(* IEC 61131-3 sources: daoli-st-library/DL_Algo (part 3) *)

(* ---- FB_DL_ThermalRampPredict.st ---- *)
(*==============================================================================
 * 组件名称 (Component)  : FB_DL_ThermalRampPredict
 * 所属子库 (Sublibrary) : DL_Algo
 * 当前版本 (Version)    : 1.0.0
 * 兼容性   (Platform)   : CODESYS 3.5+ / TwinCAT 3 / 汇川 InoProShop / 施耐德 Machine Expert
 *                         仅依赖 Standard.library（R_TRIG / ABS / MIN / MAX）与库内时间换算内核
 *                         FC_DL_TimeToLrealSec / FC_DL_LrealSecToTime，零厂商私有库
 * 功能描述 (Function)   : 一阶热模型预测与前馈。模型 dT/dt = 〔u·K − (T − Tamb)〕/ tau，本件不驱 u，
 *                         而以「满功率模型斜率」作参考，用实测斜率在线修正时间常数 tau：
 *                         ① tRemain：据当前温度、目标温度与实测斜率外推到目标所需剩余时间；
 *                         ② fFfBias：进入目标前 fLeadBand 带内按接近程度线性加大「减功率量」，
 *                         抑制热惯性造成的超调（前馈偏移，非闭环）；
 *                         ③ tau 在线修正：实测斜率与模型斜率偏差持续超阈值时按 ±5% 微调，
 *                         并钳在〔tTauMin, tTauMax〕，防单次扰动把模型带偏。
 * 分工声明 (Scope)      : 与 `FB_DL_DryingOvenZone` / `FB_DL_CvdTempRamp`（分区控温与温度曲线
 *                         执行）分工 —— 本件**只出预测与前馈偏置**，不闭环、不持曲线、不下发
 *                         加热指令；曲线执行与闭环属主为上列两件。
 * 接口     (Interface)  : 输入 fTempC 当前温度、fTargetC 目标温度、fAmbC 环境温度、fGainK 稳态
 *                         增益、tTau 时间常数、tTauMin / tTauMax 修正上下限、fLeadBand 前馈起始带、
 *                         fFfBiasMax 前馈偏置上限、fSlopeDevMax 斜率偏差阈值、tTaskPeriod 任务周期、
 *                         bEnable 使能、bReset 复位；输出 tRemain 剩余时间（无趋势时为哨兵）、
 *                         bNoTrend 无趋势标志、fFfBias 前馈减功率量、fTauUsed 当前使用的时间常数、
 *                         eState / eCause / bError / nErrId。
 * 边界     (Boundary)   : ① 组态闸：tTau <= T#0S、tTauMin <= T#0S、tTauMax <= tTauMin、fGainK <= 0.0、
 *                         fLeadBand <= 0.0、fFfBiasMax <= 0.0、fSlopeDevMax < 0.0、tTaskPeriod <= T#0S
 *                         或任一浮点引脚 NaN → 故障锁存（每个参与判据的引脚都在闸内，R151）；
 *                         ② tRemain 计算防除零：当实测斜率绝对值 <= DL_SLOPE_EPS 时**不返回 T#0S**
 *                         （T#0S 会被上层读成「马上就到」），而返回哨兵 DL_TIME_INF 并置 bNoTrend；
 *                         ③ 前馈偏置双侧钳位〔0.0, fFfBiasMax〕，禁单侧钳位；
 *                         ④ 非有限输入 → 故障闸，输出侧 tRemain 哨兵、fFfBias 0（安全侧）；
 *                         ⑤ R_TRIG 一枚段 0 无条件周期刷新；⑥ 故障相迁出唯一路径 = bReset 上升沿；
 *                         ⑦ 零全局耦合（无 GVL / 无物理地址）。
 * 遗留假设 (Assumption) : 【R95 三句声明】① 代理值 = 引脚 tTaskPeriod，用于把逐拍温差换算成 °C/s；
 *                         ② 覆盖范围 = 任务周期 10 ms ~ 2 s 的周期任务；③ 覆盖不到的区间
 *                         （< 10 ms 的高速任务或超载抖动任务）由调用方负责：此时斜率噪声偏大，
 *                         tau 修正应经 bEnable 关断，仅使用 fFfBias 前馈。
 * 解除式   (Release)    : bReset 上升沿 ∧ 组态合法 ∧ 非无趋势（NOT bNoTrend，当拍量）。
 *                         自证可满足（终审两式 1）：bNoTrend 由当拍斜率派生，温度一旦真实变化
 *                         斜率即非零，标志必落假；解除式不含计时器输出与锁存量比较，无恒假因子。
 * 码表     (Codes)      : 16#0002_03B3 故障级：热模型预测故障总码（组态非法 / 输入非有限 / 非法
 *                         相位），锁存至 bReset 上升沿，归因由 eCause 承载（R190 单件单总码）；
 *                         16#0002_04B6 信息级：无趋势（斜率近似为 0，剩余时间输出哨兵）。
 *                         加码反证（R90）：无趋势时 tRemain 是哨兵常量、fFfBias 仍有效，若只靠
 *                         「tRemain = 86400 s」判断，上层无法区分「真的还要一天」与「算不出来」，
 *                         故须立一码（bNoTrend 只是布尔位，不进报警台账）。
 *                         码段说明：0002 段故障子带 03xx / 信息子带 04xx，本件取 03B3 / 04B6
 *                         （源码实扫该两槽为空，续接同子带已用最大值，未回填碎片孔洞）。
 * 编译门槛 (Build Gate) : 本件委托 FC_DL_TimeToLrealSec 与 FC_DL_LrealSecToTime（内部转调平台
 *                         内建 TIME_TO_LREAL / LREAL_TO_TIME），交付门槛：须在 CODESYS / TwinCAT 3 /
 *                         InoProShop 三平台各编译验证一次。
 * 开源溯源 (Origin)     : 道莅自研 clean-room（参考一阶热模型与时间常数在线修正参数域，
 *                         零代码行复制；t2-1-lgf 技术子族）
 * 修订历史 (Revision)   : 2026-11-19  v1.0.0  R45 首版（批次 2 · 序号 9）
 *==============================================================================*)

TYPE E_DL_TrpState :
(
    eIdle  := 0,     // 失能待使能 / Idle, disabled
    eRun   := 10,    // 预测运行 / Predicting in run
    eFault := 90     // 故障锁存相 / Fault latched phase
);
END_TYPE

TYPE E_DL_TrpCause :
(
    eNone       := 0,   // 无故障成因 / No cause
    eCfgIllegal := 1,   // 组态非法 / Illegal configuration
    eNonFinite  := 2,   // 输入非有限 / Non-finite input
    ePhaseBad   := 3    // 非法相位兜底 / Illegal phase fallback
);
END_TYPE

FUNCTION_BLOCK FB_DL_ThermalRampPredict
VAR_INPUT
    fTempC        : REAL := 25.0;       // 当前温度 [°C] / Current temperature [degC]
    fTargetC      : REAL := 80.0;       // 目标温度 [°C] / Target temperature [degC]
    fAmbC         : REAL := 25.0;       // 环境温度 [°C] / Ambient temperature [degC]
    fGainK        : REAL := 55.0;       // 稳态增益（满功率温升上界），域 > 0.0 [°C] / Steady-state gain, domain > 0.0 [degC]
    tTau          : TIME := T#120S;     // 时间常数初值，域 > T#0S [ms] / Initial time constant, domain > T#0S [ms]
    tTauMin       : TIME := T#20S;      // 修正下限，域 > T#0S 且 < tTauMax [ms] / Correction lower bound [ms]
    tTauMax       : TIME := T#900S;     // 修正上限，域 > tTauMin [ms] / Correction upper bound [ms]
    fLeadBand     : REAL := 10.0;       // 前馈起始带（距目标多近开始减功率），域 > 0.0 [°C] / Lead band, domain > 0.0 [degC]
    fFfBiasMax    : REAL := 60.0;       // 前馈减功率量上限，域 > 0.0 [%] / Feed-forward bias ceiling, domain > 0.0 [%]
    fSlopeDevMax  : REAL := 0.05;       // 斜率偏差阈值（相对值），域 >= 0.0 [p.u.] / Slope deviation threshold [p.u.]
    tTaskPeriod   : TIME := T#100MS;    // 调用任务周期（代理值，见头注释遗留假设），域 > T#0S [ms] / Task period proxy [ms]
    bEnable       : BOOL := TRUE;       // 预测使能 [-] / Prediction enable
    bReset        : BOOL := FALSE;      // 复位命令，上升沿清故障 [-] / Reset command, rising edge clears fault
END_VAR
VAR_OUTPUT
    tRemain       : TIME;               // 剩余时间（无趋势时输出哨兵 24 h） [ms] / Remaining time, sentinel 24 h when no trend [ms]
    bNoTrend      : BOOL;               // 无趋势标志（斜率近似 0） [-] / No-trend flag
    fFfBias       : REAL;               // 前馈减功率量（双侧钳位后） [%] / Feed-forward power reduction, clamped [%]
    fTauUsed      : REAL;               // 当前使用的时间常数（在线修正后） [s] / Time constant in use after correction [s]
    eState        : E_DL_TrpState;      // 状态出口，段 6 单点映射 / State outlet
    eCause        : E_DL_TrpCause;      // 故障成因出口（R190 归因唯一） / Fault cause outlet
    bError        : BOOL;               // 故障锁存标志 [-] / Fault latch flag
    nErrId        : UDINT;              // 事件码，0 = 无事件 / Event code, 0 = no event
END_VAR
VAR
    _eState       : E_DL_TrpState := E_DL_TrpState.eIdle;   // 内部相位（CASE 唯一写入目标） / Internal phase
    _eCause       : E_DL_TrpCause := E_DL_TrpCause.eNone;   // 故障成因锁存（锁存量） / Latched cause
    rtReset       : R_TRIG;             // 复位沿实例，段 0 无条件调用 / Reset edge
    _fTsSec       : LREAL;              // 任务周期秒数（当拍量） [s] / Task period in seconds
    _fTauSec      : LREAL;              // 时间常数秒数（当拍量，取自修正后的 tTau） [s] / Time constant in seconds
    _fTempPrev    : REAL;               // 上拍温度快照（锁存量） [°C] / Previous-scan temperature snapshot
    _fSlopeMeas   : LREAL;              // 实测斜率（当拍量） [°C/s] / Measured slope [degC/s]
    _fSlopeModel  : LREAL;              // 满功率模型斜率（当拍量） [°C/s] / Full-power model slope [degC/s]
    _fDeltaT      : REAL;               // 目标 − 当前温差 [°C] / Target minus current temperature [degC]
    _fRemSec      : LREAL;              // 剩余时间秒数（转换前） [s] / Remaining seconds before conversion
    _fTauUsedSec  : LREAL;              // 在线修正后的时间常数（锁存量） [s] / Corrected time constant, latched
    _nDevRun      : INT;                // 斜率偏差持续计数（锁存量） [拍] / Slope deviation persistence counter, latched
    _uConvErrT    : UDINT;              // 周期换算错误码（当拍量） [-] / Period conversion error code
    _uConvErrU    : UDINT;              // 时间常数换算错误码（当拍量） [-] / Tau conversion error code
    _uConvErrR    : UDINT;              // 剩余时间换算错误码（当拍量） [-] / Remaining-time conversion error code
    _bConvErrT    : BOOL;               // 周期换算故障位（当拍量） [-] / Period conversion fault flag
    _bConvErrU    : BOOL;               // 时间常数换算故障位（当拍量） [-] / Tau conversion fault flag
    _bConvErrR    : BOOL;               // 剩余时间换算故障位（当拍量） [-] / Remaining-time conversion fault flag
    _bConvValidT  : BOOL;               // 周期换算有效位（当拍量） [-] / Period conversion valid flag
    _bConvValidU  : BOOL;               // 时间常数换算有效位（当拍量） [-] / Tau conversion valid flag
    _bConvValidR  : BOOL;               // 剩余时间换算有效位（当拍量） [-] / Remaining-time conversion valid flag
    _bInit        : BOOL;               // 首拍初始化完成位（锁存量） [-] / First-scan init done
    _bNonFin      : BOOL;               // 输入非有限当拍量 [-] / Non-finite input this scan
    _bCfgBad      : BOOL;               // 组态非法当拍量 [-] / Illegal configuration
    _bFault       : BOOL;               // 故障锁存位（锁存量） / Latched fault bit
    _uFault       : UDINT;              // 故障码锁存（锁存量） / Latched fault code
    _uInfo        : UDINT;              // 信息码，每拍重算 / Info code, recomputed each scan
END_VAR
VAR CONSTANT
    DL_FLOAT_EPS  : LREAL := 1.0E-6;    // 浮点判零容差 [无量纲] / Float epsilon for zero tests
    DL_SLOPE_EPS  : LREAL := 1.0E-4;    // 斜率判零容差（低于此判无趋势） [°C/s] / Slope epsilon, below means no trend [degC/s]
    DL_TIME_INF   : LREAL := 86400.0;   // 「无趋势」哨兵秒数（24 h，远离任何真实剩余时间） [s] / No-trend sentinel seconds, 24 h [s]
    DL_TAU_STEP   : LREAL := 1.05;      // 时间常数单次修正倍率 [-] / Time constant correction factor per adjustment
    DL_DEV_MAX    : INT := 10;          // 斜率偏差持续拍数门限 [拍] / Slope deviation persistence limit [scan]
END_VAR

(* —— 段 0：当拍判据派生 + 沿实例无条件周期刷新 —— *)
_fTsSec := FC_DL_TimeToLrealSec(tIn := tTaskPeriod, eErr => _uConvErrT, bError => _bConvErrT, bValid => _bConvValidT);   // 周期换算（R140 委托） / Period conversion
_fTauSec := FC_DL_TimeToLrealSec(tIn := tTau, eErr => _uConvErrU, bError => _bConvErrU, bValid => _bConvValidU);         // 时间常数换算 / Tau conversion
_bNonFin := (fTempC <> fTempC) OR (fTargetC <> fTargetC) OR (fAmbC <> fAmbC) OR (fGainK <> fGainK)    // NaN 自反判（判等禁令唯一例外） / NaN self-reflexive tests
         OR (fLeadBand <> fLeadBand) OR (fFfBiasMax <> fFfBiasMax) OR (fSlopeDevMax <> fSlopeDevMax); // 前馈参数 NaN 判 / Feed-forward parameter NaN tests
_bCfgBad := (tTau <= T#0S) OR (tTauMin <= T#0S) OR (tTauMax <= tTauMin) OR (tTaskPeriod <= T#0S)     // 时间类组态闸 / Time config gates
            OR (fGainK <= 0.0) OR (fLeadBand <= 0.0) OR (fFfBiasMax <= 0.0) OR (fSlopeDevMax < 0.0)   // 浮点域闸（R151 全覆盖） / Float domain gates
            OR (_uConvErrT <> 16#0000_0000) OR (_uConvErrU <> 16#0000_0000);                          // 换算错误并入闸 / Conversion errors folded in
rtReset(CLK := bReset);                                                                              // 复位沿，每拍必调（R228A） / Reset edge

(* —— 段 1：单拍量预清零（锁存量与快照量不入清单，R107） —— *)
_uInfo   := 16#0000_0000;          // 信息码每拍重算 / Info recomputed every scan
bNoTrend := FALSE;                 // 无趋势标志每拍预清 / No-trend flag preset
nErrId   := 16#0000_0000;          // 事件码缺省无事件 / Event code default none
bError   := FALSE;                 // 故障标志每拍预清，故障分支同拍置位（R45 配对） / Flag preset
fFfBias  := 0.0;                   // 前馈偏置缺省 0（安全侧：不减功率） / Bias default 0, safe side

(* —— 段 2：复位沿 + 组态域闸 + 非有限闸 —— *)
IF rtReset.Q THEN                                                        // 当拍复位沿 / current-scan reset edge
    _bFault := FALSE;                                                    // 清故障锁存位（锁存量） / Clear fault latch
    _uFault := 16#0000_0000;                                             // 清故障锁存码（锁存量） / Clear latched code
    _eCause := E_DL_TrpCause.eNone;                                      // 清成因（锁存量） / Clear latched cause
    IF _eState = E_DL_TrpState.eFault THEN
        _eState := E_DL_TrpState.eIdle;                                  // 故障相迁出唯一路径 / Sole exit from fault phase
    END_IF
END_IF
IF _bCfgBad THEN                                                         // 组态域闸 / Configuration gate
    _uFault := 16#0002_03B3;                                             // 故障级：热模型预测故障总码 / Fault-level: prediction fault code
    _bFault := TRUE;
    bError  := TRUE;                                                     // 故障标志同拍置位（R45 配对） / Error flag set same scan
    _eCause := E_DL_TrpCause.eCfgIllegal;                                // 归因：组态非法 / Cause: illegal configuration
END_IF
IF (NOT _bFault) AND _bNonFin THEN                                       // 输入非有限 / Non-finite input
    _uFault := 16#0002_03B3;
    _bFault := TRUE;
    bError  := TRUE;
    _eCause := E_DL_TrpCause.eNonFinite;                                 // 归因：非有限 / Cause: non-finite
END_IF

(* —— 段 3：时间常数初始化（首拍取初值并钳在修正域内） —— *)
IF NOT _bInit THEN
    IF _fTauSec < FC_DL_TimeToLrealSec(tIn := tTauMin) THEN              // 初值低于下限即钳入域内 / Clamp initial value into domain
        _fTauUsedSec := FC_DL_TimeToLrealSec(tIn := tTauMin);
    ELSIF _fTauSec > FC_DL_TimeToLrealSec(tIn := tTauMax) THEN
        _fTauUsedSec := FC_DL_TimeToLrealSec(tIn := tTauMax);
    ELSE
        _fTauUsedSec := _fTauSec;
    END_IF
    _fTempPrev := fTempC;                                                // 温度快照初始化 / Initialize temperature snapshot
    _bInit := TRUE;                                                      // 初始化完成 / Init done
END_IF

(* —— 段 4：斜率测量、模型斜率与时间常数在线修正（仅无故障且使能） —— *)
IF (NOT _bFault) AND bEnable THEN
    IF _fTsSec > DL_FLOAT_EPS THEN                                       // 除零前置判 / Divide-by-zero guard
        _fSlopeMeas := REAL_TO_LREAL(fTempC - _fTempPrev) / _fTsSec;      // 实测斜率 [°C/s] / Measured slope
    ELSE
        _fSlopeMeas := 0.0;                                              // 周期退化时置 0（组态闸已拦，防御纵深） / Degenerate period
    END_IF
    IF _fTauUsedSec > DL_FLOAT_EPS THEN                                  // 除零前置判 / Divide-by-zero guard
        _fSlopeModel := REAL_TO_LREAL(fGainK - (fTempC - fAmbC)) / _fTauUsedSec;   // 满功率模型斜率 / Full-power model slope
    ELSE
        _fSlopeModel := 0.0;                                             // 退化兜底 / Degenerate guard
    END_IF
    IF ABS(_fSlopeModel) > DL_SLOPE_EPS THEN                             // 相对偏差需有非零参照 / Relative deviation needs a non-zero reference
        IF ABS((_fSlopeMeas - _fSlopeModel) / _fSlopeModel) > fSlopeDevMax THEN
            IF _nDevRun < DL_DEV_MAX THEN
                _nDevRun := _nDevRun + 1;                                // 偏差持续计数 / Deviation persistence count
            END_IF
        ELSE
            _nDevRun := 0;                                               // 回到阈值内即清零 / Reset inside threshold
        END_IF
    ELSE
        _nDevRun := 0;
    END_IF
    IF _nDevRun >= DL_DEV_MAX THEN                                       // 偏差持续：按符号微调时间常数 / Sustained deviation, adjust tau by sign
        IF _fSlopeMeas < _fSlopeModel THEN                               // 实测偏慢 → 时间常数变大 / Slower than model, tau up
            _fTauUsedSec := MIN(_fTauUsedSec * DL_TAU_STEP, FC_DL_TimeToLrealSec(tIn := tTauMax));
        ELSE
            _fTauUsedSec := MAX(_fTauUsedSec / DL_TAU_STEP, FC_DL_TimeToLrealSec(tIn := tTauMin));
        END_IF
        _nDevRun := 0;                                                   // 修正后计数清零 / Reset after correction
    END_IF
END_IF

(* —— 段 5：剩余时间预测（防除零；无趋势输出哨兵而非 T#0S） —— *)
IF (NOT _bFault) AND bEnable THEN
    _fDeltaT := fTargetC - fTempC;                                       // 剩余温差 / Remaining temperature difference
    IF ABS(_fSlopeMeas) <= DL_SLOPE_EPS THEN                             // 斜率近似 0：不得输出 T#0S 冒充「马上到」 / Slope near zero, never emit T#0S
        bNoTrend := TRUE;                                                // 无趋势标志 / No-trend flag
        _fRemSec := DL_TIME_INF;                                         // 哨兵秒数 / Sentinel seconds
        _uInfo := 16#0002_04B6;                                          // 信息级：无趋势留痕 / Info: no trend recorded
    ELSE
        _fRemSec := REAL_TO_LREAL(_fDeltaT) / _fSlopeMeas;               // 线性外推剩余时间 / Linear extrapolation
        IF _fRemSec < 0.0 THEN                                           // 已越过目标（过冲在恢复）：剩余判 0 而非负数 / Already past target
            _fRemSec := 0.0;
        END_IF
        IF _fRemSec > DL_TIME_INF THEN                                   // 上界兜底防 TIME 溢出 / Upper bound guard
            _fRemSec := DL_TIME_INF;
        END_IF
    END_IF
    tRemain := FC_DL_LrealSecToTime(fSec := _fRemSec, eErr => _uConvErrR, bError => _bConvErrR, bValid => _bConvValidR);   // 委托时间换算 / Delegate conversion
ELSE
    tRemain := FC_DL_LrealSecToTime(fSec := DL_TIME_INF);                // 非运行相输出哨兵（不宣称「马上到」） / Sentinel outside run phase
END_IF

(* —— 段 6：前馈偏置（进入 fLeadBand 带内线性加大减功率量，双侧钳位） —— *)
IF (NOT _bFault) AND bEnable THEN
    IF ABS(_fDeltaT) < fLeadBand THEN                                    // 进入前馈带 / Inside lead band
        fFfBias := fFfBiasMax * (1.0 - (ABS(_fDeltaT) / fLeadBand));      // 越接近目标减得越多 / More reduction as target nears
    ELSE
        fFfBias := 0.0;                                                  // 带外不减功率 / No reduction outside band
    END_IF
    IF fFfBias > fFfBiasMax THEN                                         // 双侧钳位（上侧） / Two-sided clamp, upper
        fFfBias := fFfBiasMax;
    END_IF
    IF fFfBias < 0.0 THEN                                                // 双侧钳位（下侧） / Two-sided clamp, lower
        fFfBias := 0.0;
    END_IF
END_IF

(* —— 段 7：温度快照更新（主体末行，跨拍纪律） —— *)
_fTempPrev := fTempC;                                                    // 温度快照（本拍末更新） / Temperature snapshot at body end

(* —— 段 8：故障解除式（R240 全当拍量） —— *)
IF rtReset.Q AND (NOT _bCfgBad) AND (NOT _bNonFin) AND (NOT bNoTrend) THEN
    _bFault := FALSE;                                                    // 清故障锁存位（锁存量） / Clear fault latch
    _uFault := 16#0000_0000;                                             // 清故障锁存码（锁存量） / Clear latched code
    _eCause := E_DL_TrpCause.eNone;                                      // 清成因（锁存量） / Clear latched cause
END_IF

(* —— 段 8A：故障锁存相位迁移闸 —— *)
IF _bFault AND (_eState <> E_DL_TrpState.eFault) THEN
    _eState := E_DL_TrpState.eFault;                                     // 锁存即入故障相 / Latch enters fault phase
END_IF

(* —— 段 9：相位机（ENUM 全成员显式标签 + ELSE 兜底，R128） —— *)
CASE _eState OF

E_DL_TrpState.eIdle:
    IF bEnable AND _bInit AND (NOT _bFault) THEN                         // 出口 1：使能且已初始化 / Enabled and initialized
        _eState := E_DL_TrpState.eRun;
    ELSIF _bFault THEN                                                   // 出口 2：故障锁存 / Fault latched
        _eState := E_DL_TrpState.eFault;
    END_IF

E_DL_TrpState.eRun:
    IF (NOT bEnable) THEN                                                // 出口 1：失能（前置消失，R98） / Disabled
        _eState := E_DL_TrpState.eIdle;
    ELSIF _bFault THEN                                                   // 出口 2：故障锁存 / Fault latched
        _eState := E_DL_TrpState.eFault;
    END_IF

E_DL_TrpState.eFault:
    ;                                                                     // 故障相：仅段 8 复位沿可迁出 / Only the reset edge leaves this phase

ELSE
    _uFault := 16#0002_03B3;                                             // 故障级：非法相位兜底（归并总码） / Illegal-phase fallback
    _bFault := TRUE;
    bError  := TRUE;
    _eCause := E_DL_TrpCause.ePhaseBad;                                  // 归因：非法相位 / Cause: illegal phase
    _eState := E_DL_TrpState.eFault;

END_CASE

(* —— 段 10：出口单点映射（名实同源；锁存码回放；故障相安全侧） —— *)
IF _bFault THEN
    tRemain  := FC_DL_LrealSecToTime(fSec := DL_TIME_INF);               // 故障相输出哨兵（不宣称短时到达） / Sentinel in fault
    bNoTrend := TRUE;                                                    // 故障相判无趋势（不给出时间承诺） / No-trend in fault
    fFfBias  := 0.0;                                                     // 故障相不减功率（不加未知偏置） / No bias in fault
    fTauUsed := LREAL_TO_REAL(_fTauUsedSec);                             // 时间常数镜像（供调试） / Tau mirror for commissioning
ELSIF NOT bEnable THEN
    fTauUsed := LREAL_TO_REAL(_fTauUsedSec);                             // 失能相仍回放时间常数（观测语义） / Tau echoed when disabled
    tRemain  := FC_DL_LrealSecToTime(fSec := DL_TIME_INF);               // 失能相哨兵 / Sentinel when disabled
    bNoTrend := TRUE;                                                    // 失能相无预测 / No prediction when disabled
ELSE
    fTauUsed := LREAL_TO_REAL(_fTauUsedSec);                             // 运行相时间常数 / Tau in run
END_IF
IF _bFault THEN
    nErrId := _uFault;                                                   // 故障锁存码回放 / Replay latched fault code
ELSE
    nErrId := _uInfo;                                                    // 信息码 / Info code
END_IF
bError := _bFault;                                                       // 故障标志与锁存同源（名实双出口，R191） / Flag from latch
eState := _eState;                                                       // 状态出口 / State outlet
eCause := _eCause;                                                       // 成因出口 / Cause outlet

END_FUNCTION_BLOCK

(* ---- FB_DL_ValveCharacteristic.st ---- *)
(*==============================================================================
 * 组件名称 (Component)  : FB_DL_ValveCharacteristic
 * 所属子库 (Sublibrary) : DL_Algo
 * 当前版本 (Version)    : 1.0.1
 * 兼容性   (Platform)   : CODESYS 3.5 / TwinCAT 3 / 汇川 InoProShop / Machine Expert
 *                         仅依赖 Standard.library（ABS / LN / SQRT / MIN / MAX / R_TRIG）
 * 功能描述 (Function)   : 把「期望流量百分比」按调节阀固有特性折算为「阀位百分比」，
 *                         支持线性 / 等百分比 / 快开三种特性，带可调比、行程上下限、
 *                         输出死区与饱和标志。现场用途：等百分比阀按线性给定会让小流量段
 *                         分辨率不足、大流量段增益过高并引起振荡；本件把特性补偿收回
 *                         PLC 侧，工艺员不再靠「凭经验把给定调弯」。
 *                         死区只压输出抖动，不改变内部限幅结果；掉使能保持上次阀位
 *                         （阀位突跳比保持更危险），阀位回零由上层安全逻辑负责。
 * 出口契约 (Exit)       : fTravel 为最终阀位给定，域为生效行程上下限之间；
 *                         bSaturated 表示输出被流量给定域、可调比下限或行程上下限任一截断；
 *                         bError 为故障级锁存，只由 2010 / 2011 / 2012 三码置位，
 *                         bReset 上升沿清故障回空闲。信息码 2001 / 2002 / 2003 每拍重算。
 * 开源溯源 (Origin)     : 来源标签 isa88-process（工艺参数域）。许可证：ISA-88 为公开标准，
 *                         无源码可复制；调节阀流量特性公式取自公开的过程控制教材定义。
 *                         借鉴点：把「特性」做成**枚举参数域**而非三个独立功能块——三种特性
 *                         共用同一套限幅、死区与状态机，拆块会产生三份重复代码，
 *                         且特性切换在配方里属于运行期行为。
 *                         clean-room 独立实现，与任何厂商阀门功能块无代码关联。
 * 码位说明 (Codes)      : 信息级 16#0002_2001（输出被下限截断）/ 2002（输出被上限截断）/
 *                         2003（死区保持）；故障级 16#0002_2010（行程配置非法）/
 *                         2011（可调比对数的二次守卫触发）/ 2012（非法特性枚举兜底）。
 *                         共 6 码，全部落在 R12 计划第 1.2 节本件码段内。
 * 依赖     (Depends)    : 无 DL_ 内部依赖；Standard.library: ABS / LN / SQRT / MAX / R_TRIG
 * 红线自检 (Redline)    : 1 ✓ 零全局变量表依赖、零外部变量声明、零物理地址
 *                         2 ✓ 纯 IEC 61131-3，无指针、无厂商库
 *                         3 ✓ 对数与开方先做域守护、可调比下限保证对数分母不为零、
 *                             行程上下限倒置直接判故障而不交换、死区比较用容差不用判等
 *                         4 ✓ 全变量中英双语同行注释
 *                         5 ✓ 三态 ENUM + CASE 全覆盖 + ELSE 兜底（2012）；特性选择亦全覆盖
 *                         6 ✓ R_TRIG 实例在 CASE 之外每拍无条件刷新
 *                         7 ✓ END_FUNCTION_BLOCK 位于文件最后有效行
 * 规格偏离留档 (Deviation):
 *   计划 3.11 节正文提到 2004 / 2005 / 2006 三个「输入钳位」码，但同计划第 1.2 节给本件
 *   只分配了 2001~2003 与 2010~2012 六个码，两者冲突。按「码位表为准、不得自创」的纪律，
 *   本实现对输入钳位采取如下归并：流量给定越界钳位并入 2001 / 2002（越界必然让输出打端点，
 *   语义与截断一致）；可调比与死区的钳位属整定参数修正，不单独置码，仅钳位后照算，
 *   并在头注释与本段注释中写明，不再占用段外码。
 * 修订历史 (Revision)   :
 *   2026-11-15  v1.0.0  首版入库（R12 · DL_Algo 工艺参数域）
 *   2026-11-15  v1.0.1  终审修复：投运与故障复位首拍不再强制阀位回行程下限
 *                       （原实现 fLast := fLoTravel 会让阀门在复位当拍直冲最小开度，
 *                       与本件「不做阀位回零、突跳比保持更危险」的契约自相矛盾）；
 *                       改为「保持上次阀位并夹到生效行程内」，同时补齐行程域的出口保证
 *============================================================================*)

(*-----------------------------------------------------------------------------
 * 枚举: E_DL_ValveCharKind（归属 DL_Algo，与本功能块同文件）
 * 含义: 调节阀固有流量特性。三种特性共用同一套限幅与死区逻辑。
 *----------------------------------------------------------------------------*)
TYPE E_DL_ValveCharKind :
(
    eLinear       := 0,    // 线性特性：阀位与流量成正比 / Linear: travel proportional to flow
    eEqualPercent := 10,   // 等百分比特性：单位阀位变化引起的流量变化与当前流量成正比 / Equal percentage
    eQuickOpen    := 20    // 快开特性：小阀位即获大流量，后段渐平 / Quick opening, fast rise then flat
);
END_TYPE

(*-----------------------------------------------------------------------------
 * 枚举: E_DL_ValveCharState（归属 DL_Algo，与本功能块同文件）
 * 含义: 特性补偿块的离散状态。
 *----------------------------------------------------------------------------*)
TYPE E_DL_ValveCharState :
(
    eIdle   := 0,     // 空闲：等待使能与行程配置校验 / Idle: waiting for enable and travel validation
    eActive := 10,    // 运行：折算特性、限幅、死区、输出 / Active: convert, clamp, deadband, publish
    eFault  := 99     // 故障：配置非法或枚举兜底，输出保持上次 / Fault: invalid config, travel held
);
END_TYPE

(*==============================================================================
 * 功能块: FB_DL_ValveCharacteristic
 * 调用约定: 每个扫描周期无条件调用一次；bEnable 为 FALSE 时阀位保持上次值。
 * 无状态泄漏: 全部状态驻留于实例私有 VAR，零全局引用，可多实例并行。
 *============================================================================*)
FUNCTION_BLOCK FB_DL_ValveCharacteristic
VAR_INPUT
    bEnable       : BOOL;                                // 使能，FALSE 时阀位保持上次输出 / Enable, holds the last travel when FALSE
    bReset        : BOOL;                                // 上升沿清故障回空闲 / Rising edge clears the fault
    fFlowCmd      : REAL := 0.0;                         // 期望流量 [百分比]，域 0~100 / Desired flow in percent, 0..100
    eChar         : E_DL_ValveCharKind := E_DL_ValveCharKind.eEqualPercent;  // 固有特性 [-] / Inherent characteristic
    fRangeability : REAL := 30.0;                        // 可调比 [-]，域 2~100，越界钳位 / Rangeability, clamped to 2..100
    fMinTravel    : REAL := 0.0;                         // 最小阀位 [百分比]，域 0~100 / Minimum travel in percent
    fMaxTravel    : REAL := 100.0;                       // 最大阀位 [百分比]，域 0~100 / Maximum travel in percent
    fDeadband     : REAL := 0.2;                         // 输出死区 [百分比]，变化小于此值保持上次 / Output deadband in percent
END_VAR
VAR_OUTPUT
    fTravel       : REAL;                                // 阀位给定 [百分比]，域 fMinTravel~fMaxTravel / Travel command in percent
    bSaturated    : BOOL;                                // 输出被上下限或可调比下限截断 TRUE / Output clamped
    bError        : BOOL;                                // 故障级锁存，仅 2010~2012 置位 / Latched fault
    uErrorId      : UDINT;                               // 事件码，0 = 无事件 / Event code, zero means none
    eState        : E_DL_ValveCharState;                 // 主状态机当前状态 / Current state
END_VAR
VAR
    fbTrigReset   : R_TRIG;                              // 复位沿，CASE 之外每拍刷新 / Reset edge, refreshed outside CASE
    ePhase        : E_DL_ValveCharState := E_DL_ValveCharState.eIdle;  // 内部状态 / Internal state
    fFlowVal      : REAL;                                // 钳位后的期望流量 [百分比] / Clamped flow command in percent
    fQ            : REAL;                                // 归一化流量 [0~1] / Normalised flow
    fR            : REAL;                                // 生效可调比 [-] / Effective rangeability
    fRaw          : REAL;                                // 未限幅的阀位 [百分比] / Unlimited travel in percent
    fLast         : REAL;                                // 上次输出阀位 [百分比] / Last travel command
    fLoTravel     : REAL;                                // 生效行程下限 [百分比] / Effective lower bound
    fHiTravel     : REAL;                                // 生效行程上限 [百分比] / Effective upper bound
    fQMin         : REAL;                                // 可调比下限对应的归一化流量 [0~1] / Normalised flow at the rangeability floor
    fDeadUse      : REAL;                                // 生效死区宽度 [百分比] / Effective deadband width
    bClampLo      : BOOL;                                // 下限截断标记 / Lower clamp flag
    bClampHi      : BOOL;                                // 上限截断标记 / Upper clamp flag
END_VAR
VAR CONSTANT
    DL_PCT_MAX    : REAL := 100.0;                       // 百分比满量程 [百分比] / Percent full scale
    DL_R_MIN      : REAL := 2.0;                         // 可调比下限 [-] / Minimum rangeability
    DL_R_MAX      : REAL := 100.0;                       // 可调比上限 [-] / Maximum rangeability
    DL_DB_MAX     : REAL := 5.0;                         // 死区宽度上限 [百分比] / Deadband ceiling in percent
    DL_EPS        : REAL := 1.0E-6;                      // 浮点判零容差 [-] / Float zero tolerance
END_VAR

(*------------------------------------------------------------------------------
 * 段 1｜复位沿每拍无条件刷新（严禁放进 CASE 内部）
 *      Reset edge refreshed unconditionally on every scan
 *-----------------------------------------------------------------------------*)
fbTrigReset(CLK := bReset);

(*------------------------------------------------------------------------------
 * 段 2｜输入调理：流量给定的域钳位，与整定参数的可调比 / 死区钳位
 *      Input conditioning: flow clamp plus rangeability and deadband clamps
 *      流量越界钳位必然把输出打到端点，语义等同截断，故并入 2001 / 2002 报码
 *      A clamped flow command drives the output to an end point, reported as 2001 / 2002
 *      可调比与死区的钳位只是整定参数修正，不单独置码，钳位后照算
 *      Rangeability and deadband clamps are tuning fixes and carry no dedicated code
 *-----------------------------------------------------------------------------*)
bClampLo  := FALSE;
bClampHi  := FALSE;
fFlowVal  := fFlowCmd;
IF NOT (fFlowVal >= 0.0) THEN
    fFlowVal := 0.0;
    bClampLo := TRUE;
ELSIF fFlowVal > DL_PCT_MAX THEN
    fFlowVal := DL_PCT_MAX;
    bClampHi := TRUE;
END_IF

fR := fRangeability;
IF NOT ((fR >= DL_R_MIN) AND (fR <= DL_R_MAX)) THEN
    IF fR > DL_R_MAX THEN
        fR := DL_R_MAX;
    ELSIF fR < DL_R_MIN THEN
        fR := DL_R_MIN;
    ELSE
        (* 非有限值：按上限处理，保证对数分母远离零 *)
        (* Non finite value: fall back to the ceiling so the logarithm stays safe *)
        fR := DL_R_MAX;
    END_IF
END_IF

fDeadUse := ABS(fDeadband);
IF NOT (fDeadUse <= DL_DB_MAX) THEN
    fDeadUse := DL_DB_MAX;
END_IF

fLoTravel := fMinTravel;
fHiTravel := fMaxTravel;

(*------------------------------------------------------------------------------
 * 段 3｜主状态机：三态全覆盖 + ELSE 兜底；掉使能只保持阀位，不推进任何相位
 *      Main state machine; a disabled block only holds the travel
 *-----------------------------------------------------------------------------*)
IF NOT bEnable THEN
    fTravel    := fLast;
    bSaturated := FALSE;
ELSE

    CASE ePhase OF
        E_DL_ValveCharState.eIdle:
            (* 行程配置校验：越界或倒置一律判故障，绝不静默交换上下限 *)
            (* Travel validation: out of range or inverted is a fault, never swapped *)
            IF NOT ((fMinTravel >= 0.0) AND (fMinTravel <= DL_PCT_MAX)) THEN
                bError   := TRUE;
                uErrorId := 16#0002_2010;
                ePhase   := E_DL_ValveCharState.eFault;
            ELSIF NOT ((fMaxTravel >= 0.0) AND (fMaxTravel <= DL_PCT_MAX)) THEN
                bError   := TRUE;
                uErrorId := 16#0002_2010;
                ePhase   := E_DL_ValveCharState.eFault;
            ELSIF fMinTravel > fMaxTravel THEN
                bError   := TRUE;
                uErrorId := 16#0002_2010;
                ePhase   := E_DL_ValveCharState.eFault;
            ELSE
                (* 投运与故障复位不强制阀位回零：保持上次阀位并夹到生效行程内 *)
                (* Commissioning and fault reset hold the last travel, clamped into the travel band *)
                fLast      := MIN(MAX(fLast, fLoTravel), fHiTravel);
                fTravel    := fLast;
                bSaturated := FALSE;
                uErrorId   := 16#0000_0000;
                ePhase     := E_DL_ValveCharState.eActive;
            END_IF

        E_DL_ValveCharState.eActive:
            (* 信息码每拍重算，故障码由 bError 锁存 *)
            (* Informational codes are recomputed every scan, faults stay latched *)
            uErrorId   := 16#0000_0000;
            bSaturated := FALSE;
            fQ         := fFlowVal / DL_PCT_MAX;

            CASE eChar OF
                E_DL_ValveCharKind.eLinear:
                    fRaw := fQ * DL_PCT_MAX;

                E_DL_ValveCharKind.eEqualPercent:
                    fQMin := 1.0 / fR;
                    IF fQ <= fQMin THEN
                        (* 低于可调比下限：阀位归零并记下限截断 *)
                        (* Below the rangeability floor: travel drops to zero *)
                        fRaw     := 0.0;
                        bClampLo := TRUE;
                    ELSE
                        IF ABS(LN(fR)) < DL_EPS THEN
                            (* 二次守卫：正常钳位下不可达，防调用方绕过钳位直接注入 *)
                            (* Second guard: unreachable after clamping, protects against bypass *)
                            bError   := TRUE;
                            uErrorId := 16#0002_2011;
                            ePhase   := E_DL_ValveCharState.eFault;
                        ELSE
                            fRaw := DL_PCT_MAX * (1.0 + LN(fQ) / LN(fR));
                        END_IF
                    END_IF

                E_DL_ValveCharKind.eQuickOpen:
                    (* 先取零下界再开方，浮点误差导致的负小数不会变成非数 *)
                    (* Clamp to zero before the square root so rounding cannot yield NaN *)
                    fRaw := DL_PCT_MAX * (1.0 - SQRT(MAX(0.0, 1.0 - fQ)));

                ELSE
                    (* 非法特性枚举：终端安全态 + 段内末码 *)
                    (* Illegal characteristic: terminal safe state with the segment last code *)
                    bError   := TRUE;
                    uErrorId := 16#0002_2012;
                    ePhase   := E_DL_ValveCharState.eFault;
            END_CASE

            IF ePhase = E_DL_ValveCharState.eActive THEN
                (* 行程限幅：夹到生效上下限，截断方向决定报哪个信息码 *)
                (* Travel clamp: report the direction together with the clamp *)
                IF fRaw < fLoTravel THEN
                    fRaw     := fLoTravel;
                    bClampLo := TRUE;
                ELSIF fRaw > fHiTravel THEN
                    fRaw     := fHiTravel;
                    bClampHi := TRUE;
                END_IF

                IF bClampLo THEN
                    bSaturated := TRUE;
                    IF uErrorId = 16#0000_0000 THEN
                        uErrorId := 16#0002_2001;
                    END_IF
                END_IF
                IF bClampHi THEN
                    bSaturated := TRUE;
                    IF uErrorId = 16#0000_0000 THEN
                        uErrorId := 16#0002_2002;
                    END_IF
                END_IF

                (* 死区：只压输出抖动，内部限幅结果保持不变，比较用容差不用判等 *)
                (* Deadband suppresses jitter only, the clamped value stays untouched *)
                IF ABS(fRaw - fLast) < fDeadUse THEN
                    fTravel := fLast;
                    IF uErrorId = 16#0000_0000 THEN
                        uErrorId := 16#0002_2003;
                    END_IF
                ELSE
                    fTravel := fRaw;
                    fLast   := fRaw;
                END_IF
            END_IF

        E_DL_ValveCharState.eFault:
            (* 故障态保持上次阀位，只认复位沿；不在故障态做任何折算 *)
            (* Fault holds the last travel and only the reset edge leaves it *)
            fTravel := fLast;
            IF fbTrigReset.Q THEN
                bError   := FALSE;
                uErrorId := 16#0000_0000;
                ePhase   := E_DL_ValveCharState.eIdle;
            END_IF

        ELSE
            (* 兜底：枚举被在线改坏或跨版本不兼容，阀位保持并等待复位 *)
            (* Fallback: hold the travel and wait for a reset *)
            bError   := TRUE;
            uErrorId := 16#0002_2012;
            fTravel  := fLast;
            ePhase   := E_DL_ValveCharState.eFault;
    END_CASE

END_IF

(*------------------------------------------------------------------------------
 * 段 4｜状态出口：内部状态镜像到出口引脚，便于 HMI 直接显示
 *      State mirror to the output pin for direct HMI display
 *-----------------------------------------------------------------------------*)
eState := ePhase;
END_FUNCTION_BLOCK

(* ---- FC_DL_AirDensityFanPower.st ---- *)
(*==============================================================================
 * 组件名称 (Component)  : FC_DL_AirDensityFanPower
 * 所属子库 (Sublibrary) : DL_Algo
 * 当前版本 (Version)    : 1.0.0
 * 兼容性 (Platform)     : CODESYS 3.5 / TwinCAT 3 / 汇川 InoProShop / Machine Expert
 *                         仅依赖纯 IEC 61131-3 标准元素，零厂商方言
 * 功能描述 (Function)   : 风机轴功率空气密度修正：P_corr = P_rated x rho/rho0，
 *                         rho 委托 FC_DL_AirDensity（湿空气理想气体内核）
 *                         本函数只做前置校验 + 钳位 + 错误码，不重写密度内核。
 * 溯源 (Origin)         : 道莅 clean-room 防御性实现
 * 本文件内含 (Contains) : TYPE E_DL_FanErr / FUNCTION FC_DL_AirDensityFanPower
 * 依赖 (Depends)        : DL_Algo/FC_DL_AirDensity
 * 红线自检 (Redline)    : 无外部全局变量、无硬件地址直引 ｜ 全变量中英双语同行注释
 *                         防除零 + 量程钳位 + 非有限值防御 ｜ 枚举成员全部显式赋值
 *                         纯函数无状态保持 ｜ 输出在每条早退路径前已赋确定值
 * 错误码表 (Codes)      : 16#0002_370B 成功
 *                         16#0002_370C 信息级 温度越界(已钳制)
 *                         16#0002_370D 信息级 湿度越界(已钳制)
 *                         16#0002_370E 信息级 压力越界(已钳制)
 *                         16#0002_370F 故障级 额定功率非法（<= 0 或非有限）
 * 修订历史 (Revision)   : 2026-11-17  v1.0.0  首版入库 · R27 · 阶段三批 1
 * 验收向量 (Acceptance) : T=20 C, RH=50%, P=101325 Pa → rho≈1.2041，
 *                         ratio≈0.9829, P_rated=10 kW → P_corr≈9.829 kW，返回 370B
 *============================================================================*)

(*-----------------------------------------------------------------------------
 * 枚举: E_DL_FanErr（归属 DL_Algo，与 FC_DL_AirDensityFanPower 同文件）
 *----------------------------------------------------------------------------*)
TYPE E_DL_FanErr :
(
    eOk          := 16#0002_370B,    // 成功 / Success
    eTempClamped := 16#0002_370C,    // 信息级：温度越界已钳制 / Info: temperature clamped
    eHumClamped  := 16#0002_370D,    // 信息级：湿度越界已钳制 / Info: humidity clamped
    ePressClamp  := 16#0002_370E,    // 信息级：压力越界已钳制 / Info: pressure clamped
    ePowerBad    := 16#0002_370F     // 故障级：额定功率非法 / Fault: illegal rated power
);
END_TYPE

(*==============================================================================
 * 函数: FC_DL_AirDensityFanPower（纯函数，无任何状态保持）
 * 调用约定: 每周期按需调用；返回值 = 计算有效标志。
 *============================================================================*)
FUNCTION FC_DL_AirDensityFanPower : BOOL
VAR_INPUT
    fTemp_C     : REAL;                // 气温 [摄氏度]，有效域 -40~60 / Air temperature [degC]
    fRelHumPct  : REAL;                // 相对湿度 [百分数]，有效域 0~100 / Relative humidity [percent]
    fPress_Pa   : REAL;                // 大气压 [帕]，有效域 6.0E4~1.1E5 / Atmospheric pressure [Pa]
    fPowerRated : REAL;                // 额定轴功率 [千瓦]，有效域 0.1~5000 / Rated shaft power [kW]
END_VAR
VAR_OUTPUT
    fPowerCorr  : REAL;                // 密度修正后轴功率 [千瓦] / Density-corrected shaft power [kW]
    eError      : E_DL_FanErr;         // 错误码 / Error code
END_VAR
VAR CONSTANT
    DL_FAN_T_MIN     : REAL := -40.0;   // 温度域下限 [摄氏度] / Temperature lower bound [degC]
    DL_FAN_T_MAX     : REAL := 60.0;    // 温度域上限 [摄氏度] / Temperature upper bound [degC]
    DL_FAN_HUM_MIN   : REAL := 0.0;     // 湿度域下限 [百分数] / Humidity lower bound [percent]
    DL_FAN_HUM_MAX   : REAL := 100.0;   // 湿度域上限 [百分数] / Humidity upper bound [percent]
    DL_FAN_P_MIN     : REAL := 6.0E4;   // 大气压域下限 [帕] / Pressure lower bound [Pa]
    DL_FAN_P_MAX     : REAL := 1.1E5;   // 大气压域上限 [帕] / Pressure upper bound [Pa]
    DL_FAN_RHO0      : REAL := 1.225;   // 标准工况空气密度 [千克每立方米] / Reference air density [kg/m3]
    DL_FAN_RATIO_MIN : REAL := 0.5;     // 密度比强制下限 [无量纲] / Forced ratio lower bound
    DL_FAN_RATIO_MAX : REAL := 1.5;     // 密度比强制上限 [无量纲] / Forced ratio upper bound
    DL_FAN_INF_MAX   : REAL := 1.0E30;  // 非有限值判定幅值上限 / Magnitude bound for finite-value check
    DL_FAN_ZERO      : REAL := 0.0;     // 零值常量，避免裸字面量 / Zero constant
END_VAR
VAR
    fTempUse  : REAL;                  // 生效温度（钳位后）[摄氏度] / Effective temperature [degC]
    fHumUse   : REAL;                  // 生效湿度（钳位后）[百分数] / Effective humidity [percent]
    fPressUse : REAL;                  // 生效大气压（钳位后）[帕] / Effective pressure [Pa]
    fRho      : LREAL;                 // 委托密度输出 [千克每立方米] / Density from the delegate [kg/m3]
    fRatio    : REAL;                  // 密度比 rho/rho0 [无量纲] / Density ratio [dimensionless]
    bNonFin   : BOOL;                  // 非有限输入汇总标志 / Non-finite input aggregate flag
END_VAR

(*------------------------------------------------------------------------------
 * 段 1｜出口默认值：任何早退路径前输出已确定（哨兵 0 功率 + 功率非法码）
 *----------------------------------------------------------------------------*)
FC_DL_AirDensityFanPower := FALSE;                   // 返回值默认无效 / return defaults to invalid
fPowerCorr := DL_FAN_ZERO;                           // 功率哨兵 0 / power sentinel zero
eError := E_DL_FanErr.ePowerBad;                     // 默认功率非法码 / default illegal-power code

(*------------------------------------------------------------------------------
 * 段 2｜非有限值闸：NaN 用自反判，溢出用幅值上限判
 *----------------------------------------------------------------------------*)
bNonFin := (fTemp_C     <> fTemp_C)     OR (ABS(fTemp_C)     > DL_FAN_INF_MAX)
        OR (fRelHumPct  <> fRelHumPct)  OR (ABS(fRelHumPct)  > DL_FAN_INF_MAX)
        OR (fPress_Pa   <> fPress_Pa)   OR (ABS(fPress_Pa)   > DL_FAN_INF_MAX)
        OR (fPowerRated <> fPowerRated) OR (ABS(fPowerRated) > DL_FAN_INF_MAX);
IF bNonFin THEN
    eError := E_DL_FanErr.ePowerBad;                 // 非有限输入并入功率非法段（同为全拒，反证句见头注）/ non-finite mapped to power band
    RETURN;
END_IF

(*------------------------------------------------------------------------------
 * 段 3｜额定功率闸：必须为正且落在可信域
 *----------------------------------------------------------------------------*)
IF (fPowerRated < 0.1) OR (fPowerRated > 5000.0) THEN
    eError := E_DL_FanErr.ePowerBad;                 // 故障级：额定功率非法 / fault: illegal rated power
    RETURN;
END_IF

(*------------------------------------------------------------------------------
 * 段 4｜三输入钳位（信息级越界码，温度→湿度→压力优先级顺序判定）
 *----------------------------------------------------------------------------*)
eError := E_DL_FanErr.eOk;                           // 预置成功 / preset success
fTempUse := fTemp_C;                                 // 温度工作副本 / temperature working copy
IF fTempUse < DL_FAN_T_MIN THEN
    fTempUse := DL_FAN_T_MIN;                        // 下限钳位 / floored
    eError := E_DL_FanErr.eTempClamped;              // 信息级：温度越界 / info: temperature clamped
ELSIF fTempUse > DL_FAN_T_MAX THEN
    fTempUse := DL_FAN_T_MAX;                        // 上限钳位 / capped
    eError := E_DL_FanErr.eTempClamped;              // 信息级：温度越界 / info: temperature clamped
END_IF
fHumUse := fRelHumPct;                               // 湿度工作副本 / humidity working copy
IF fHumUse < DL_FAN_HUM_MIN THEN
    fHumUse := DL_FAN_HUM_MIN;                       // 下限钳位 / floored
    IF eError = E_DL_FanErr.eOk THEN
        eError := E_DL_FanErr.eHumClamped;           // 信息级：湿度越界（不覆盖前序码）/ info: humidity clamped
    END_IF
ELSIF fHumUse > DL_FAN_HUM_MAX THEN
    fHumUse := DL_FAN_HUM_MAX;                       // 上限钳位 / capped
    IF eError = E_DL_FanErr.eOk THEN
        eError := E_DL_FanErr.eHumClamped;           // 信息级：湿度越界（不覆盖前序码）/ info: humidity clamped
    END_IF
END_IF
fPressUse := fPress_Pa;                              // 压力工作副本 / pressure working copy
IF fPressUse < DL_FAN_P_MIN THEN
    fPressUse := DL_FAN_P_MIN;                       // 下限钳位 / floored
    IF eError = E_DL_FanErr.eOk THEN
        eError := E_DL_FanErr.ePressClamp;           // 信息级：压力越界（不覆盖前序码）/ info: pressure clamped
    END_IF
ELSIF fPressUse > DL_FAN_P_MAX THEN
    fPressUse := DL_FAN_P_MAX;                       // 上限钳位 / capped
    IF eError = E_DL_FanErr.eOk THEN
        eError := E_DL_FanErr.ePressClamp;           // 信息级：压力越界（不覆盖前序码）/ info: pressure clamped
    END_IF
END_IF

(*------------------------------------------------------------------------------
 * 段 5｜委托密度（FC_DL_AirDensity 湿空气内核）
 *----------------------------------------------------------------------------*)
fRho := FC_DL_AirDensity(fTempC := REAL_TO_LREAL(fTempUse), fPressPa := REAL_TO_LREAL(fPressUse), fRh := REAL_TO_LREAL(fHumUse));   // 密度委托 [千克每立方米] / density via delegate
IF (fRho <> fRho) OR (ABS(fRho) > REAL_TO_LREAL(DL_FAN_INF_MAX)) OR (fRho <= LREAL#1.0E-9) THEN
    eError := E_DL_FanErr.ePowerBad;                 // 委托输出不可信：按功率非法全拒处置（反证句：输出同为哨兵+无效）/ unusable delegate output
    fPowerCorr := DL_FAN_ZERO;                       // 功率哨兵 / power sentinel
    FC_DL_AirDensityFanPower := FALSE;               // 返回无效 / return invalid
    RETURN;
END_IF

(*------------------------------------------------------------------------------
 * 段 6｜密度比计算与强制钳位 [0.5, 1.5]：除子 rho0 为常量非零
 *----------------------------------------------------------------------------*)
fRatio := LREAL_TO_REAL(fRho) / DL_FAN_RHO0;         // 密度比 [无量纲] / density ratio [dimensionless]
IF fRatio < DL_FAN_RATIO_MIN THEN
    fRatio := DL_FAN_RATIO_MIN;                      // 比率强制下限（防过修）/ forced ratio floor
ELSIF fRatio > DL_FAN_RATIO_MAX THEN
    fRatio := DL_FAN_RATIO_MAX;                      // 比率强制上限（防过修）/ forced ratio ceiling
END_IF

(*------------------------------------------------------------------------------
 * 段 7｜功率修正与出口（P = P_rated x ratio）
 *----------------------------------------------------------------------------*)
fPowerCorr := fPowerRated * fRatio;                  // 修正功率 [千瓦] / corrected power [kW]
IF fPowerCorr > DL_FAN_INF_MAX THEN
    fPowerCorr := DL_FAN_INF_MAX;                    // 溢出钳位防护 / overflow clamp guard
END_IF
IF fPowerCorr < DL_FAN_ZERO THEN
    fPowerCorr := DL_FAN_ZERO;                       // 下限防护 / floor guard
END_IF
FC_DL_AirDensityFanPower := TRUE;                    // 计算有效 / computation valid
RETURN;
END_FUNCTION

(* ---- FC_DL_BiquadCoeff.st ---- *)
(*
  ==================================================================
  组件名 Component  : FC_DL_BiquadCoeff
  分类   Category   : DL_Algo
  前缀   Naming     : FC_DL_ ｜ b/n/u/f/t/e/st 类型前缀制（R265）
  码位   Code ID    : 16#0002_373D / 373E（故障级）
  版本   Version    : 1.0.0
  复杂度 Complexity  : 中
  功能   Purpose    : 二阶节五系数生成器（低通 / 高通 / 带通 / 陷波四型，归一化
                      a0 = 1 口径），为 FB_DL_BiquadFilter / FB_DL_BiquadCascade
                      提供下发系数，闭合「设计 → 下发」链。
  开源溯源 Origin    : 公开公式 clean-room，参考 RBJ Audio EQ Cookbook 类公开二阶节
                      设计公式（biquad coefficient 公式为公开领域知识，分类与公式
                      借鉴，零代码复制），本件实现、闸门与码位 100% 自有。
  许可证 License    : MIT
  参考   Reference  : IEC 61131-3:2013 §6.6 算术运算符；RBJ Audio EQ Cookbook 公开
                      二阶节设计公式（w0 = 2π·f0/Fs，alpha = sin(w0)/(2Q)）
  平台   Platform   : 纯 IEC 61131-3（FOR / CASE / 四则 / SIN / COS），三平台通用
  依赖   Depends    : 仅 Standard.library（SIN / COS 属标准内建）
  分工声明 Split     : FB_DL_NotchFilter（陷波一体机：内算内滤）/ FB_DL_SecondOrder
                      Filter（巴特沃斯二阶：内算内滤）为内算型；本件只产系数**不下发
                      执行**，与两个内算型互引，现场自行组合（R216）。
  归属 Ownership     : E_DL_BiquadType 属主为本文件（全库唯一定义，R264）；引用件
                      只引用不重声明。
  ------------------------------------------------------------------
  边界 Boundary     :
                      一 域闸全量枚举（R272）：fFs ≤ 0、fF0 ≤ 0 或 ≥ 0.45×fFs
                         （奈奎斯特闸）、fQ 越域 [0.1, 20.0]、任一非有限 → 五系数
                         全 0 + 故障码 373D + 三件套 + RETURN 结构早退；
                      二 枚举越域（CASE ELSE）：落 373D 同码处置——反证句（R90）：
                         枚举非法与域闸失败的出口组合完全同形（五系数全 0、bValid =
                         FALSE），无法由输出区分，按 R90 不另立码；
                      三 归一化除子 a0 = 1 + alpha：alpha > 0 结构性成立（fF0 > 0
                         已证 → w0 ∈ (0, 0.9π) → sin(w0) > 0 → alpha > 0 → a0 > 1），
                         另设 ABS(a0) < 1.0E-9 闸（码 373E）作平台数值兜底；
                      四 中间量常量提级：2π、0.45 与 Q 域界全部 VAR CONSTANT，
                         禁魔法数；
                      五 Jury 一致性声明：本件产出的系数建议由 FB_DL_BiquadFilter /
                         BiquadCascade 的 Jury 三条件闸复验；两闸口径一致
                         （|a2|<1 ∧ 1+a1+a2>0 ∧ 1−a1+a2>0，返修 R2 固化判据）；
                      六 结果复检非有限 → 三件套兜底（R258）；
                      七 纯函数：无记忆量、无定时器、无边沿实例，每调用重算；
                      八 无全局、无外部变量、无物理地址、无指针。
  错误码 Codes      :
    16#0002_373D【故障级】域闸失败（fFs / fF0 / fQ 越域或任一非有限，或类型枚举
                         非法，五系数全 0）
    16#0002_373E【故障级】归一化分母近零（ABS(a0) < 1.0E-9）或结果复检非有限
                         （后者理论上不可达的兜底分支，出口组合同形，R90 不另立）
  码位反证 Note     :
    373D 与 373E 不可合并：373D 出口五系数全 0 且未进入计算，373E 出口同样全 0 但
    已进入计算，两者处置人不同（组态工程师调参数 / 数值平台问题），且 373E 仅在
    理论上不可达路径出现，按 R90 分立两码（场景可由码值唯一还原）。
  验收 Acceptance   :
    算法已证（脚本）：未跑 ｜ 编译器已证（三平台）：未跑
    V1 fFs = 1000, fF0 = 100, fQ = 0.7071 低通（巴特沃斯）→ b0 ≈ 0.06745、
       b1 ≈ 0.1349、b2 ≈ 0.06745、a1 ≈ −1.1430、a2 ≈ 0.4128（公开设计值）
    V2 同参高通 → 系数为低通镜像（b0 / b2 互换语义，b1 取负）
    V3 fF0 = 0.46×fFs → 奈奎斯特闸故障早退；V4 fQ = 0 → 故障早退
    V5 fFs = 0 → 故障早退；V6 陷波型 fF0 = 50, fFs = 1000, fQ = 5 → 在 50Hz
       处增益 ≈ 0（定性向量）；V7 fQ = 25 → 越域故障早退
  修订记录 Revision  :
    2026-11-21  v1.0.0  R63 首版（批 2 · 序号 6）
  ==================================================================
*)
TYPE E_DL_BiquadType :
(
    eLowPass  := 0, // 低通：通带以下通过，截止频率以上衰减 / the low pass type passing below the cutoff
    eHighPass := 1, // 高通：截止频率以上通过，以下衰减 / the high pass type passing above the cutoff
    eBandPass := 2, // 带通：中心频率附近通过（0 dB 峰值增益口径）/ the band pass type passing around the center with a zero dB peak gain
    eNotch    := 3  // 陷波：中心频率处深衰减（挖槽）/ the notch type with a deep attenuation at the center
);
END_TYPE

FUNCTION FC_DL_BiquadCoeff : BOOL
VAR_INPUT
    eType   : E_DL_BiquadType := E_DL_BiquadType.eLowPass; // 滤波器类型 [-] / the filter type
    fFs     : LREAL := 1000.0; // 采样频率 [赫兹]，须 > 0 / the sampling frequency, must be positive
    fF0     : LREAL := 100.0;  // 中心 / 截止频率 [赫兹]，0 < fF0 < 0.45×fFs / the center or cutoff frequency below the Nyquist guard
    fQ      : LREAL := 0.7071; // 品质因数 [−]，域 [0.1, 20.0] / the quality factor inside its domain
END_VAR
VAR_OUTPUT
    fB0     : LREAL := 0.0; // 归一化前向系数 b0 [−]，a0 = 1 口径 / the normalized feed forward coefficient b0
    fB1     : LREAL := 0.0; // 归一化前向系数 b1 [−] / the normalized feed forward coefficient b1
    fB2     : LREAL := 0.0; // 归一化前向系数 b2 [−] / the normalized feed forward coefficient b2
    fA1     : LREAL := 0.0; // 归一化反馈系数 a1 [−] / the normalized feedback coefficient a1
    fA2     : LREAL := 0.0; // 归一化反馈系数 a2 [−] / the normalized feedback coefficient a2
    bValid  : BOOL := FALSE; // 结果可用 [-] / the result usable flag
    eErr    : UDINT := 16#0000_0000; // 错误码，0 = 正常 / the error code, zero is ok
    bError  : BOOL := FALSE; // 故障标志（故障级码同拍置位，R45 配对）/ the fault flag raised with a fault level code
END_VAR
VAR
    fW0     : LREAL := 0.0; // 数字角频率 w0 = 2π·f0/Fs [弧度] / the digital angular frequency
    fCosW0  : LREAL := 0.0; // cos(w0) 中间量 [−] / the cosine intermediate
    fSinW0  : LREAL := 0.0; // sin(w0) 中间量 [−] / the sine intermediate
    fAlpha  : LREAL := 0.0; // 阻尼因子 alpha = sin(w0)/(2Q) [−]，除子 2Q 已证 > 0 / the damping factor with the proven divisor
    fA0     : LREAL := 0.0; // 归一化前分母 a0 = 1 + alpha [−] / the pre normalization denominator
    fB0Raw  : LREAL := 0.0; // 未归一化 b0 暂存 [−] / the raw b0 in staging
    fB1Raw  : LREAL := 0.0; // 未归一化 b1 暂存 [−] / the raw b1 in staging
    fB2Raw  : LREAL := 0.0; // 未归一化 b2 暂存 [−] / the raw b2 in staging
    fA1Raw  : LREAL := 0.0; // 未归一化 a1 暂存 [−] / the raw a1 in staging
    fA2Raw  : LREAL := 0.0; // 未归一化 a2 暂存 [−] / the raw a2 in staging
    fNyq    : LREAL := 0.0; // 奈奎斯特闸限 0.45×fFs [赫兹] / the Nyquist guard value
END_VAR  // R64 结构补齐：VAR 段缺失的 END_VAR（门禁机械修复）
VAR CONSTANT
    DL_BQC_2PI   : LREAL := 6.283185307179586; // 2π 常量（LREAL 精度字面量，R55）/ the two pi constant at LREAL precision
    DL_BQC_NYQ   : LREAL := 0.45;   // 奈奎斯特闸系数 [−]（0.45×fFs）/ the Nyquist guard fraction
    DL_BQC_QMIN  : LREAL := 0.1;    // 品质因数下界 [−] / the quality factor floor
    DL_BQC_QMAX  : LREAL := 20.0;   // 品质因数上界 [−] / the quality factor ceiling
    DL_BQC_DENEPS: LREAL := 1.0E-9; // 归一化分母近零门限 [−] / the near zero denominator threshold
    DL_BQC_TWO   : LREAL := 2.0;    // 实数二常量 [−]（阻尼因子除子）/ the real two constant
    DL_BQC_ZERO  : LREAL := 0.0;    // 实数零常量 [−] / the real zero constant
    DL_BQC_ONE   : LREAL := 1.0;    // 实数一常量 [−] / the real one constant
    DL_BQC_HALF  : LREAL := 0.5;    // 实数半常量 [−] / the real half constant
END_VAR

// 段 1｜返回值与全部出口预置安全值（R45 四段式第一段：五系数全 0）/ segment 1, the preset of the return and every outlet
FC_DL_BiquadCoeff := FALSE; // 返回值预置假 / preset the return false
fB0 := DL_BQC_ZERO; // 系数 b0 预置零 [−] / preset the coefficient b0 zero
fB1 := DL_BQC_ZERO; // 系数 b1 预置零 [−] / preset the coefficient b1 zero
fB2 := DL_BQC_ZERO; // 系数 b2 预置零 [−] / preset the coefficient b2 zero
fA1 := DL_BQC_ZERO; // 系数 a1 预置零 [−] / preset the coefficient a1 zero
fA2 := DL_BQC_ZERO; // 系数 a2 预置零 [−] / preset the coefficient a2 zero
bValid := FALSE; // 可用标志预置假 / preset the validity false
eErr := 16#0000_0000; // 错误码预置正常 / preset the code to ok
bError := FALSE; // 故障标志预置假 / preset the error flag false
fW0 := DL_BQC_ZERO; // 角频率预置零 [弧度] / preset the angular frequency zero
fCosW0 := DL_BQC_ZERO; // 余弦预置零 [−] / preset the cosine zero
fSinW0 := DL_BQC_ZERO; // 正弦预置零 [−] / preset the sine zero
fAlpha := DL_BQC_ZERO; // 阻尼因子预置零 [−] / preset the damping zero
fA0 := DL_BQC_ZERO; // 分母预置零 [−] / preset the denominator zero
fB0Raw := DL_BQC_ZERO; // 原始 b0 预置零 [−] / preset the raw b0 zero
fB1Raw := DL_BQC_ZERO; // 原始 b1 预置零 [−] / preset the raw b1 zero
fB2Raw := DL_BQC_ZERO; // 原始 b2 预置零 [−] / preset the raw b2 zero
fA1Raw := DL_BQC_ZERO; // 原始 a1 预置零 [−] / preset the raw a1 zero
fA2Raw := DL_BQC_ZERO; // 原始 a2 预置零 [−] / preset the raw a2 zero
fNyq := DL_BQC_ZERO; // 奈奎斯特闸限预置零 [赫兹] / preset the Nyquist guard zero

// 段 2｜域闸全量枚举（边界一，R272：fFs / fF0 / fQ 逐个点名 + 非有限双判）/ segment 2, the full domain gate naming every real pin
fNyq := DL_BQC_NYQ * fFs; // 奈奎斯特闸限（fFs 非有限时乘积亦非有限，闸随后命中）[赫兹] / the Nyquist guard, a non finite sampling frequency lands non finite and the gate catches it
IF (fFs <> fFs) OR ((fFs - fFs) <> (fFs - fFs)) OR (fFs <= DL_BQC_ZERO)
OR (fF0 <> fF0) OR ((fF0 - fF0) <> (fF0 - fF0)) OR (fF0 <= DL_BQC_ZERO) OR (fF0 >= fNyq)
OR (fQ <> fQ) OR ((fQ - fQ) <> (fQ - fQ)) OR (fQ < DL_BQC_QMIN) OR (fQ > DL_BQC_QMAX) THEN // 域闸失败 / a domain gate failure
    eErr := 16#0002_373D; // 故障级：域闸失败 / fault grade, a domain gate failure
    bError := TRUE; // 同拍置故障标志（R45 配对）/ raise the fault flag on the same scan
    bValid := FALSE; // 结果不可用 / the result is not usable
    RETURN; // 结构早退：五系数已预置全 0，计算段不可达 / the structural early exit with all five coefficients preset to zero
END_IF

// 段 3｜中间量计算（除子 fFs 已证 > 0、2Q 已证 > 0.2）/ segment 3, the intermediates
fW0 := (DL_BQC_2PI * fF0) / fFs; // 数字角频率 [弧度]，除子已证 > 0 / the angular frequency with the proven divisor
fCosW0 := COS(fW0); // cos(w0) [−] / the cosine
fSinW0 := SIN(fW0); // sin(w0) [−] / the sine
fAlpha := fSinW0 / (DL_BQC_TWO * fQ); // 阻尼因子 [−]，除子已证 > 0 / the damping factor with the proven divisor
fA0 := DL_BQC_ONE + fAlpha; // 归一化前分母 [−]，结构性 > 1（边界三证明）/ the pre normalization denominator structurally above one

// 段 4｜四型未归一化系数（CASE 必带 ELSE 兜底，边界二）/ segment 4, the four raw coefficient families
CASE eType OF
    E_DL_BiquadType.eLowPass: // 低通 / the low pass family
        fB0Raw := (DL_BQC_ONE - fCosW0) * DL_BQC_HALF; // b0 = (1−cos w0)/2 [−] / the raw b0
        fB1Raw := DL_BQC_ONE - fCosW0; // b1 = 1−cos w0 [−] / the raw b1
        fB2Raw := (DL_BQC_ONE - fCosW0) * DL_BQC_HALF; // b2 = (1−cos w0)/2 [−] / the raw b2
        fA1Raw := -DL_BQC_TWO * fCosW0; // a1 = −2·cos w0 [−] / the raw a1
        fA2Raw := DL_BQC_ONE - fAlpha; // a2 = 1−alpha [−] / the raw a2
    E_DL_BiquadType.eHighPass: // 高通 / the high pass family
        fB0Raw := (DL_BQC_ONE + fCosW0) * DL_BQC_HALF; // b0 = (1+cos w0)/2 [−] / the raw b0
        fB1Raw := -(DL_BQC_ONE + fCosW0); // b1 = −(1+cos w0) [−] / the raw b1
        fB2Raw := (DL_BQC_ONE + fCosW0) * DL_BQC_HALF; // b2 = (1+cos w0)/2 [−] / the raw b2
        fA1Raw := -DL_BQC_TWO * fCosW0; // a1 = −2·cos w0 [−] / the raw a1
        fA2Raw := DL_BQC_ONE - fAlpha; // a2 = 1−alpha [−] / the raw a2
    E_DL_BiquadType.eBandPass: // 带通（0 dB 峰值增益口径）/ the band pass family
        fB0Raw := fAlpha; // b0 = alpha [−] / the raw b0
        fB1Raw := DL_BQC_ZERO; // b1 = 0 [−] / the raw b1
        fB2Raw := -fAlpha; // b2 = −alpha [−] / the raw b2
        fA1Raw := -DL_BQC_TWO * fCosW0; // a1 = −2·cos w0 [−] / the raw a1
        fA2Raw := DL_BQC_ONE - fAlpha; // a2 = 1−alpha [−] / the raw a2
    E_DL_BiquadType.eNotch: // 陷波 / the notch family
        fB0Raw := DL_BQC_ONE; // b0 = 1 [−] / the raw b0
        fB1Raw := -DL_BQC_TWO * fCosW0; // b1 = −2·cos w0 [−] / the raw b1
        fB2Raw := DL_BQC_ONE; // b2 = 1 [−] / the raw b2
        fA1Raw := -DL_BQC_TWO * fCosW0; // a1 = −2·cos w0 [−] / the raw a1
        fA2Raw := DL_BQC_ONE - fAlpha; // a2 = 1−alpha [−] / the raw a2
    ELSE // 枚举非法：落 373D 同码（反证句见码表，出口与域闸失败同形）/ an illegal enumeration under the same code
        eErr := 16#0002_373D; // 故障级：类型枚举非法（归入域闸族）/ fault grade, the type enumeration is illegal in the gate family
        bError := TRUE; // 同拍置故障标志（R45 配对）/ raise the fault flag on the same scan
        bValid := FALSE; // 结果不可用 / the result is not usable
        RETURN; // 早退，五系数保持预置全 0 / early return with the preset zeros
END_CASE

// 段 5｜归一化除子闸与系数归一（边界三，禁除零）/ segment 5, the normalization with the denominator guard
IF ABS(fA0) < DL_BQC_DENEPS THEN // 分母近零（理论不可达的平台数值兜底）/ a near zero denominator, a platform numerical fallback
    eErr := 16#0002_373E; // 故障级：归一化分母近零 / fault grade, the normalization denominator is near zero
    bError := TRUE; // 同拍置故障标志（R45 配对）/ raise the fault flag on the same scan
    bValid := FALSE; // 结果不可用 / the result is not usable
    RETURN; // 早退，五系数保持全 0 / early return with the zeros
END_IF
fB0 := fB0Raw / fA0; // 归一化 b0 [−]，除子已证 ≥ 门限 / the normalized b0
fB1 := fB1Raw / fA0; // 归一化 b1 [−] / the normalized b1
fB2 := fB2Raw / fA0; // 归一化 b2 [−] / the normalized b2
fA1 := fA1Raw / fA0; // 归一化 a1 [−] / the normalized a1
fA2 := fA2Raw / fA0; // 归一化 a2 [−] / the normalized a2

// 段 6｜结果复检兜底（三件套，R258；与 373E 同码，反证见码表）/ segment 6, the result recheck with the three part fallback
IF (fB0 <> fB0) OR ((fB0 - fB0) <> (fB0 - fB0))
OR (fB1 <> fB1) OR ((fB1 - fB1) <> (fB1 - fB1))
OR (fB2 <> fB2) OR ((fB2 - fB2) <> (fB2 - fB2))
OR (fA1 <> fA1) OR ((fA1 - fA1) <> (fA1 - fA1))
OR (fA2 <> fA2) OR ((fA2 - fA2) <> (fA2 - fA2)) THEN // 任一系数非有限（理论上不可达，防御保留）/ any non finite coefficient, unreachable by theory
    fB0 := DL_BQC_ZERO; // 系数 b0 兜底归零 [−] / the bottom line zero
    fB1 := DL_BQC_ZERO; // 系数 b1 兜底归零 [−] / the bottom line zero
    fB2 := DL_BQC_ZERO; // 系数 b2 兜底归零 [−] / the bottom line zero
    fA1 := DL_BQC_ZERO; // 系数 a1 兜底归零 [−] / the bottom line zero
    fA2 := DL_BQC_ZERO; // 系数 a2 兜底归零 [−] / the bottom line zero
    eErr := 16#0002_373E; // 故障级：结果非有限（同族一码）/ fault grade under the same family code
    bError := TRUE; // 置故障标志（R45 配对）/ raise the fault flag
    bValid := FALSE; // 结果不可用 / the result is not usable
    RETURN; // 早退 / early return
END_IF

// 段 7｜统一出口 / segment 7, the unified outlet
bValid := TRUE; // 结果可用 / the result is usable
FC_DL_BiquadCoeff := TRUE; // 返回成功 / return success
END_FUNCTION

(* ---- FC_DL_GasFlowSqrt.st ---- *)
(*==============================================================================
 * 组件名称 (Component)  : FC_DL_GasFlowSqrt
 * 所属子库 (Sublibrary) : DL_Algo
 * 当前版本 (Version)    : 1.0.0
 * 兼容性 (Platform)     : CODESYS 3.5 / TwinCAT 3 / 汇川 InoProShop / Machine Expert
 *                         仅依赖纯 IEC 61131-3 标准元素，零厂商方言
 * 功能描述 (Function)   : 特气差压流量开方换算：前置校验 → 补偿系数钳位 →
 *                         委托 FC_DL_NthRoot(2) 开方 → 委托 FC_DL_FlowCompensate
 *                         做温压补偿内核（固定参考工况口径）→ 量程换算 → 上限钳制。
 *                         本函数不重写任何开方/补偿数学内核（T0 红线）。
 * 溯源 (Origin)         : 道莅 clean-room 防御性实现
 * 本文件内含 (Contains) : TYPE E_DL_FlowErr / FUNCTION FC_DL_GasFlowSqrt
 * 依赖 (Depends)        : DL_MathData/FC_DL_NthRoot、DL_Algo/FC_DL_FlowCompensate
 * 红线自检 (Redline)    : 无外部全局变量、无硬件地址直引 ｜ 全变量中英双语同行注释
 *                         防除零 + 量程钳位 + 非有限值防御 ｜ 枚举成员全部显式赋值
 *                         纯函数无状态保持 ｜ 输出在每条早退路径前已赋确定值
 * 错误码表 (Codes)      : 16#0002_3706 成功
 *                         16#0002_3707 故障级 密度非法（<= 0 或非有限）
 *                         16#0002_3708 故障级 差压为负
 *                         16#0002_3709 信息级 补偿系数越界(已钳制)
 *                         16#0002_370A 故障级 结果溢出或委托失败
 * 修订历史 (Revision)   : 2026-11-17  v1.0.0  首版入库 · R27 · 阶段三批 1
 * 验收向量 (Acceptance) : dp=25 kPa, rho=2.0, comp=1.0, scale=100 slm
 *                         → sqrt(25/100)*1.0*100 = 50 slm，返回 3706
 *============================================================================*)

(*-----------------------------------------------------------------------------
 * 枚举: E_DL_FlowErr（归属 DL_Algo，与 FC_DL_GasFlowSqrt 同文件）
 *----------------------------------------------------------------------------*)
TYPE E_DL_FlowErr :
(
    eOk           := 16#0002_3706,   // 成功 / Success
    eDensityBad   := 16#0002_3707,   // 故障级：密度非法（<= 0 或非有限）/ Fault: illegal density
    eDiffPressNeg := 16#0002_3708,   // 故障级：差压为负 / Fault: negative differential pressure
    eCompClamped  := 16#0002_3709,   // 信息级：补偿系数越界已钳制 / Info: compensation factor clamped
    eResultOver   := 16#0002_370A    // 故障级：结果溢出或委托失败 / Fault: result overflow or delegate failure
);
END_TYPE

(*==============================================================================
 * 函数: FC_DL_GasFlowSqrt（纯函数，无任何状态保持）
 * 调用约定: 每周期按需调用；返回值 = 计算有效标志。
 * 口径说明: 差压满刻度取 DL_GSF_DP_FULL（100 kPa），根号归一化后乘补偿系数
 *           与满量程；补偿内核（温压链）委托 FC_DL_FlowCompensate 固定参考
 *           工况执行，外部 fCompFactor 为调用方注入的合成补偿比。
 *============================================================================*)
FUNCTION FC_DL_GasFlowSqrt : BOOL
VAR_INPUT
    fDiffPress   : REAL;               // 差压 [千帕]，有效域 0~100 / Differential pressure [kPa]
    fGasDensity  : REAL;               // 工况密度 [千克每立方米]，有效域 0.01~20 / Gas density at operating condition [kg/m3]
    fCompFactor  : REAL;               // 温压补偿系数 [无量纲]，有效域 0.5~2.0 / Compensation factor [dimensionless]
    fScaleMax    : REAL;               // 流量满量程 [标准升每分钟]，须 > 0 / Full-scale flow [slm]
END_VAR
VAR_OUTPUT
    fFlowSlm     : REAL;               // 流量 [标准升每分钟] / Flow [slm]
    eError       : E_DL_FlowErr;       // 错误码 / Error code
END_VAR
VAR CONSTANT
    DL_GSF_DP_FULL  : REAL := 100.0;   // 差压满刻度 [千帕] / Full-scale differential pressure [kPa]
    DL_GSF_COMP_MIN : REAL := 0.5;     // 补偿系数下限 [无量纲] / Compensation factor lower bound
    DL_GSF_COMP_MAX : REAL := 2.0;     // 补偿系数上限 [无量纲] / Compensation factor upper bound
    DL_GSF_T_REF    : REAL := 20.0;    // 委托补偿参考温度 [摄氏度] / Delegate compensation reference temperature [degC]
    DL_GSF_INF_MAX  : REAL := 1.0E30;  // 非有限值判定幅值上限 / Magnitude bound for finite-value check
    DL_GSF_ZERO     : REAL := 0.0;     // 零值常量，避免裸字面量 / Zero constant
    DL_GSF_RHO_MIN  : REAL := 0.01;    // 密度可信下限 [千克每立方米] / Density trust lower bound [kg/m3]
    DL_GSF_RHO_MAX  : REAL := 20.0;    // 密度可信上限 [千克每立方米] / Density trust upper bound [kg/m3]
END_VAR
VAR
    fCompUse   : REAL;                 // 生效补偿系数（钳位后）[无量纲] / Effective compensation factor
    fRootVal   : LREAL;                // 委托开方输出 [无量纲合成] / Delegate square-root output
    bRootOk    : BOOL;                 // 委托开方有效标志 / Delegate root validity flag
    fCompFlow  : REAL;                 // 委托补偿后的流量基值 [标准升每分钟] / Delegate-compensated flow base [slm]
    uCompErr   : UDINT;                // 委托补偿错误码（0 = 无错）/ Delegate compensation error id
    bCompRange : BOOL;                 // 委托补偿域内标志 / Delegate in-range flag
    bNonFin    : BOOL;                 // 非有限输入汇总标志 / Non-finite input aggregate flag
END_VAR

(*------------------------------------------------------------------------------
 * 段 1｜出口默认值：任何早退路径前输出已确定（哨兵 0 流量 + 输入无效码）
 *----------------------------------------------------------------------------*)
FC_DL_GasFlowSqrt := FALSE;                          // 返回值默认无效 / return defaults to invalid
fFlowSlm := DL_GSF_ZERO;                             // 流量哨兵 0 / flow sentinel zero
eError := E_DL_FlowErr.eDensityBad;                  // 默认密度非法码 / default illegal-density code

(*------------------------------------------------------------------------------
 * 段 2｜非有限值闸：NaN 用自反判，溢出用幅值上限判
 *----------------------------------------------------------------------------*)
bNonFin := (fDiffPress  <> fDiffPress)  OR (ABS(fDiffPress)  > DL_GSF_INF_MAX)
        OR (fGasDensity <> fGasDensity) OR (ABS(fGasDensity) > DL_GSF_INF_MAX)
        OR (fCompFactor <> fCompFactor) OR (ABS(fCompFactor) > DL_GSF_INF_MAX)
        OR (fScaleMax   <> fScaleMax)   OR (ABS(fScaleMax)   > DL_GSF_INF_MAX);
IF bNonFin THEN
    eError := E_DL_FlowErr.eDensityBad;              // 非有限输入并入密度非法段（反证句见文件头修订）/ non-finite mapped to density band
    RETURN;
END_IF

(*------------------------------------------------------------------------------
 * 段 3｜符号与配置闸：密度可信域、差压非负、满量程为正
 *----------------------------------------------------------------------------*)
IF (fGasDensity < DL_GSF_RHO_MIN) OR (fGasDensity > DL_GSF_RHO_MAX) OR (fScaleMax <= DL_GSF_ZERO) THEN
    eError := E_DL_FlowErr.eDensityBad;              // 故障级：密度非法（含满量程非法并入，反证句：同为全拒）/ fault: illegal density
    RETURN;
END_IF
IF fDiffPress < DL_GSF_ZERO THEN
    eError := E_DL_FlowErr.eDiffPressNeg;            // 故障级：差压为负 / fault: negative dp
    RETURN;
END_IF

(*------------------------------------------------------------------------------
 * 段 4｜补偿系数钳位（信息级越界码）
 *----------------------------------------------------------------------------*)
eError := E_DL_FlowErr.eOk;                          // 预置成功 / preset success
fCompUse := fCompFactor;                             // 补偿系数工作副本 / compensation working copy
IF fCompUse < DL_GSF_COMP_MIN THEN
    fCompUse := DL_GSF_COMP_MIN;                     // 下限钳位 / floored
    eError := E_DL_FlowErr.eCompClamped;             // 信息级：补偿系数越界 / info: factor clamped
ELSIF fCompUse > DL_GSF_COMP_MAX THEN
    fCompUse := DL_GSF_COMP_MAX;                     // 上限钳位 / capped
    eError := E_DL_FlowErr.eCompClamped;             // 信息级：补偿系数越界 / info: factor clamped
END_IF

(*------------------------------------------------------------------------------
 * 段 5｜委托开方（FC_DL_NthRoot(2)）：差压满刻度归一化后的根号值
 *----------------------------------------------------------------------------*)
fRootVal := FC_DL_NthRoot(fValue := REAL_TO_LREAL(fDiffPress / DL_GSF_DP_FULL), nRoot := 2, bValid => bRootOk);   // 根号委托（除子 100 为常量非零）/ root via delegate
IF (NOT bRootOk) OR (fRootVal <> fRootVal) OR (ABS(fRootVal) > REAL_TO_LREAL(DL_GSF_INF_MAX)) THEN
    eError := E_DL_FlowErr.eResultOver;              // 故障级：委托失败 / fault: delegate failure
    FC_DL_GasFlowSqrt := FALSE;                      // 返回无效 / return invalid
    RETURN;
END_IF

(*------------------------------------------------------------------------------
 * 段 6｜委托温压补偿内核（FC_DL_FlowCompensate 固定参考工况口径，满量程换算）
 *----------------------------------------------------------------------------*)
fCompFlow := FC_DL_FlowCompensate(fFlowActual := LREAL_TO_REAL(fRootVal) * fScaleMax * fCompUse,   // 委托入口流量 [标准升每分钟] / delegate input flow [slm]
                                  fPressGauge := DL_GSF_ZERO,                                     // 固定参考表压 [千帕] / fixed reference gauge pressure [kPa]
                                  fTempC := DL_GSF_T_REF,                                         // 固定参考温度 [摄氏度] / fixed reference temperature [degC]
                                  bEnableSqRt := FALSE,                                           // 开方已在段 5 委托完成 / root already delegated
                                  uErrorId => uCompErr, bInRange => bCompRange);                  // 委托出口 / delegate outputs
IF (uCompErr <> 0) OR (fCompFlow <> fCompFlow) OR (ABS(fCompFlow) > DL_GSF_INF_MAX) THEN
    eError := E_DL_FlowErr.eResultOver;              // 故障级：补偿委托失败或结果溢出 / fault: delegate failure or overflow
    fFlowSlm := DL_GSF_ZERO;                         // 流量哨兵 / flow sentinel
    FC_DL_GasFlowSqrt := FALSE;                      // 返回无效 / return invalid
    RETURN;
END_IF

(*------------------------------------------------------------------------------
 * 段 7｜上限钳制与出口
 *----------------------------------------------------------------------------*)
fFlowSlm := fCompFlow;                               // 流量输出 [标准升每分钟] / flow output [slm]
IF fFlowSlm > fScaleMax THEN
    fFlowSlm := fScaleMax;                           // 满量程钳制 / clamped to full scale
END_IF
IF fFlowSlm < DL_GSF_ZERO THEN
    fFlowSlm := DL_GSF_ZERO;                         // 下限防护（禁止伪负流量）/ floor guard
END_IF
FC_DL_GasFlowSqrt := TRUE;                           // 计算有效 / computation valid
RETURN;
END_FUNCTION

(* ---- FC_DL_HeatExchangerLmtd.st ---- *)
(*
  FC_DL_HeatExchangerLmtd  —  换热器对数平均温差 + ε-NTU 效能 / Heat exchanger LMTD and effectiveness
  分类 Category : DL_Algo
  码位 Code     : 16#02_3_84
  版本 Version  : 1.0.0
  来源 Source   : t2-1-lgf-technology — IEC 61131-3 标准语义的道莅防御性实现
  溯源 Origin   : clean-room 实现，LMTD/ε-NTU 公开传热语义，未复制任何源码行
  功能 Function : 1) 按流向布置（逆流/并流/1-2 程）取端差 ΔT1/ΔT2，LMTD = (ΔT1−ΔT2)/LN(ΔT1/ΔT2)；
                  2) 1-2 程乘 F 修正系数（Kern 公式，R≈1 走极限分支）；
                  3) 效能 ε：NTU = U·A/(m·cp)，Cr 由端差能量平衡反推（Cr = MIN(r, 1/r)，r = ΔTh/ΔTc）；
                  4) 热侧换热量 fQkw = m·cp·(T_h,in − T_h,out) / 1000。
  边界 Boundary : ① ΔT1 与 ΔT2 符号相反 → bTempCross := TRUE 置故障码（温度交叉，物理不可能）；
                  ② 任一 ΔT <= 0 判无效置码；|ΔT1−ΔT2| < 1E-3 K 走退化分支改算术平均（禁 LN(1) 除零）；
                  ③ fMassFlowHotKgS <= 0 / fCpHotJkgK <= 0 / fAreaM2 <= 0 防除零判组态错；
                  ④ fUwPerM2K <= 0 时仅输出 fLmtdK，fEpsilon := 0 并置「UA 未组态」信息码（Q 亦不输出）；
                  ⑤ F 修正分支：P >= 1 或 P·R >= 1 判退化（端点温度重合），1-2 程不输出效能；
                  ⑥ 解除式自证：bTempCross/bDegenerate 每调用重算，条件消失即自动解除（无锁存）。
  依赖 Depends  : 仅 Standard.library（LN/EXP/SQRT/ABS/MIN/MAX）；枚举 E_DL_FlowArrangement 随本件发布
  码表 Error codes（本件格 02_3_84，子码步进 +0x100）:
    16#0002_0184 信息级：UA 未组态（U <= 0），仅输出 LMTD，效能/热量不输出
    16#0002_0284 故障级：温度交叉（ΔT1 与 ΔT2 符号相反）或任一端差 <= 0
    16#0002_0384 故障级：组态非法（m <= 0 / cp <= 0 / A <= 0）
    16#0002_0484 信息级：端差退化分支（|ΔT1−ΔT2| < 1E-3 K，改算术平均）
    16#0002_0584 故障级：1-2 程 F 修正域退化（P >= 1 或 P·R >= 1，端点重合）

  修订历史 Revision :
    2026-11-18  v1.0.0  R38 首版
*)

TYPE E_DL_FlowArrangement :
(
    eCounter         := 0,   // 逆流 / Counter flow
    eParallel        := 1,   // 并流 / Parallel flow
    eOneShellTwoTube := 2    // 1-2 程（壳侧 1 程，管侧 2 程）/ One shell pass, two tube passes
);
END_TYPE

FUNCTION FC_DL_HeatExchangerLmtd : BOOL
VAR_INPUT
    fHotInC        : REAL;                        // 热侧进口温度 [°C] / Hot inlet temperature
    fHotOutC       : REAL;                        // 热侧出口温度 [°C] / Hot outlet temperature
    fColdInC       : REAL;                        // 冷侧进口温度 [°C] / Cold inlet temperature
    fColdOutC      : REAL;                        // 冷侧出口温度 [°C] / Cold outlet temperature
    eFlowType      : E_DL_FlowArrangement;        // 流向布置 / Flow arrangement
    fAreaM2        : REAL;                        // 换热面积 [m²]，域 > 0 / Heat transfer area
    fUwPerM2K      : REAL;                        // 总传热系数 U [W/(m²·K)]，<= 0 = 未组态 / Overall U coefficient
    fMassFlowHotKgS: REAL;                        // 热侧质量流量 [kg/s]，域 > 0 / Hot side mass flow
    fCpHotJkgK     : REAL;                        // 热侧比热 [J/(kg·K)]，域 > 0 / Hot side specific heat
END_VAR
VAR_OUTPUT
    fLmtdK         : REAL;                        // 对数平均温差 [K] / Log mean temperature difference
    fEpsilon       : REAL;                        // 效能 [无量纲 0..1] / Effectiveness
    fQkw           : REAL;                        // 热侧换热量 [kW] / Heat duty
    bTempCross     : BOOL;                        // 温度交叉标志 / Temperature cross flag
    bDegenerate    : BOOL;                        // 端差退化标志（改算术平均）/ Degenerate-end-difference flag
    nErrId         : UDINT;                       // 事件码，0 = 无事件 / Event code, 0 = none
END_VAR
VAR
    rDt1, rDt2     : LREAL;                       // 两端差 [K] / Terminal differences
    rLmtd, rNum    : LREAL;                       // LMTD 与分子暂存 / LMTD and numerator scratch
    rCph, rRatio   : LREAL;                       // 热侧热容流率/端差比 / Hot capacity rate, delta ratio
    rNtu, rCr      : LREAL;                       // NTU 与热容比 / NTU and capacity ratio
    rR, rP, rX, rF : LREAL;                       // 1-2 程修正中间量 / One-shell-two-tube F correction scratch
    rLnArg         : LREAL;                       // 对数自变量暂存 / Logarithm argument scratch
END_VAR
VAR CONSTANT
    rDtEps   : LREAL := 1.0E-3;   // 端差退化阈值 [K] / End-difference degeneracy threshold
    rEpsMin  : LREAL := 1.0E-6;   // R≈1 判据阈值 / R near-unity threshold
    rZeroMin : LREAL := 1.0E-12; // 近零判据通用阈值 / Generic near-zero threshold
END_VAR

(* —— 段 1：输出缺省与组态闸（纯函数，每调用重算） —— *)
fLmtdK := 0.0;  fEpsilon := 0.0;  fQkw := 0.0;    // 输出缺省 0
bTempCross := FALSE;  bDegenerate := FALSE;       // 判据标志缺省
nErrId := 16#0000_0000;                           // 事件码缺省无事件
FC_DL_HeatExchangerLmtd := FALSE;                 // 返回值缺省失败

IF (LREAL(fMassFlowHotKgS) <= rZeroMin) OR (LREAL(fCpHotJkgK) <= rZeroMin)
   OR (LREAL(fAreaM2) <= rZeroMin) THEN
    nErrId := 16#0002_0384;                       // 故障级：组态非法（防除零）
    RETURN;
END_IF

(* —— 段 2：按布置取端差（ΔT 均取「热侧 − 冷侧」，符号即物理方向） —— *)
CASE eFlowType OF

E_DL_FlowArrangement.eCounter:
    rDt1 := LREAL(fHotInC)  - LREAL(fColdOutC);   // 逆流：进口端差 = 热 进 − 冷 出
    rDt2 := LREAL(fHotOutC) - LREAL(fColdInC);    // 逆流：出口端差 = 热 出 − 冷 进

E_DL_FlowArrangement.eParallel:
    rDt1 := LREAL(fHotInC)  - LREAL(fColdInC);    // 并流：进口端差 = 热 进 − 冷 进
    rDt2 := LREAL(fHotOutC) - LREAL(fColdOutC);   // 并流：出口端差 = 热 出 − 冷 出

E_DL_FlowArrangement.eOneShellTwoTube:
    rDt1 := LREAL(fHotInC)  - LREAL(fColdOutC);   // 1-2 程：按逆流端点取端差（F 修正承载差异）
    rDt2 := LREAL(fHotOutC) - LREAL(fColdInC);

ELSE
    nErrId := 16#0002_0384;                       // 未知布置并入组态错兜底
    RETURN;

END_CASE

(* —— 段 3：温度交叉与端差有效性判据 —— *)
IF (rDt1 > 0.0) <> (rDt2 > 0.0) THEN
    bTempCross := TRUE;                           // 端差符号相反：温度交叉（物理不可能）
END_IF
IF (rDt1 <= 0.0) OR (rDt2 <= 0.0) OR bTempCross THEN
    nErrId := 16#0002_0284;                       // 故障级：温度交叉或端差 <= 0
    RETURN;                                       // 不输出 LMTD
END_IF

(* —— 段 4：LMTD（退化分支改算术平均，禁 LN(1) 除零） —— *)
IF ABS(rDt1 - rDt2) < rDtEps THEN
    rLmtd := (rDt1 + rDt2) / 2.0;                 // 退化分支：算术平均（规格强制）
    bDegenerate := TRUE;                          // 退化标志
    nErrId := 16#0002_0484;                       // 信息级：端差退化分支
ELSE
    rNum := rDt1 - rDt2;                          // 分子（已闸 |·| >= 1E-3）
    rLmtd := rNum / LN(rDt1 / rDt2);              // 对数平均（分母 LN(ΔT1/ΔT2) 与分子同号，非零）
END_IF
fLmtdK := REAL(rLmtd);

(* —— 段 5：UA 未组态短路（仅输出 LMTD） —— *)
IF LREAL(fUwPerM2K) <= rZeroMin THEN
    nErrId := 16#0002_0184;                       // 信息级：UA 未组态
    FC_DL_HeatExchangerLmtd := TRUE;              // LMTD 已有效输出
    RETURN;                                       // fEpsilon/fQkw 维持 0
END_IF

(* —— 段 6：ε-NTU 效能（Cr 由端差能量平衡反推） —— *)
rCph := LREAL(fMassFlowHotKgS) * LREAL(fCpHotJkgK);               // 热侧热容流率 [W/K]
rNtu := LREAL(fUwPerM2K) * LREAL(fAreaM2) / rCph;                 // NTU = U·A/(m·cp)，分母已闸
rRatio := rDt1 / MAX(rDt2, rDtEps);                               // r = ΔTh/ΔTc（冷端差用作 ΔTc 已闸 > 0）
rCr := MIN(rRatio, 1.0 / rRatio);                                 // Cr = Cmin/Cmax ∈ [0,1]，防除零（rRatio > 0）
IF ABS(rCr - 1.0) < rEpsMin THEN
    fEpsilon := REAL(rNtu / (1.0 + rNtu));                        // Cr = 1 极限：ε = NTU/(1+NTU)
ELSIF eFlowType = E_DL_FlowArrangement.eParallel THEN
    fEpsilon := REAL((1.0 - EXP(-rNtu * (1.0 + rCr))) / (1.0 + rCr));  // 并流效能式
ELSE
    fEpsilon := REAL((1.0 - EXP(-rNtu * (1.0 - rCr)))
              / (1.0 - rCr * EXP(-rNtu * (1.0 - rCr))));          // 逆流/1-2 程效能式
END_IF

IF eFlowType = E_DL_FlowArrangement.eOneShellTwoTube THEN
    rR := rRatio;                                                 // R = ΔTh/ΔTc
    rP := 1.0 - rDt2 / MAX(LREAL(fHotInC) - LREAL(fColdInC), rDtEps);  // P = (Tco−Tci)/(Thi−Tci)
    IF (rP <= 0.0) OR (rP >= 1.0) OR (rP * rR >= 1.0) THEN
        nErrId := 16#0002_0584;                                   // 故障级：F 修正域退化（端点重合）
        RETURN;
    END_IF
    rX := SQRT(rR * rR + 1.0);                                    // X = sqrt(R²+1)
    IF ABS(rR - 1.0) < rEpsMin THEN
        rLnArg := (2.0 - rP * (2.0 - rX)) / (2.0 - rP * (2.0 + rX));  // R = 1 极限分支的对数自变量
        rF := (rX * rP / (1.0 - rP)) / LN(rLnArg);                // R = 1 极限：F = X·P/((1−P)·ln(·))
    ELSE
        rLnArg := (1.0 - rP) / (1.0 - rP * rR);                   // 通用分支第一对数自变量（已闸 > 0）
        rF := (rX / (rR - 1.0)) * LN(rLnArg)
            / LN((2.0 - rP * (rR + 1.0 - rX)) / (2.0 - rP * (rR + 1.0 + rX)));  // Kern 通用式
    END_IF
    fEpsilon := REAL(MIN(MAX(LREAL(fEpsilon) * rF, 0.0), 1.0));   // 效能乘 F 修正并钳 0..1
END_IF

(* —— 段 7：热侧换热量与出口 —— *)
fQkw := REAL(rCph * (LREAL(fHotInC) - LREAL(fHotOutC)) / 1000.0); // Q = m·cp·ΔTh [kW]
fEpsilon := REAL(MIN(MAX(LREAL(fEpsilon), 0.0), 1.0));            // 效能钳 0..1
FC_DL_HeatExchangerLmtd := TRUE;                                  // 计算有效

END_FUNCTION

(* ---- FC_DL_HumidityRatioCalc.st ---- *)
//==============================================================================
// 函数：FC_DL_HumidityRatioCalc ｜ 中文名称：含湿量计算（焓湿图族拆分②）
// 所属子库：DL_Algo ｜ 版本：v1.0.1 ｜ 兼容：CODESYS V3.5+ / TwinCAT 3 / 汇川 InoProShop
// 功能描述：由干球温度 + 露点或相对湿度求含湿量 W = 0.621945·p_v/(p−p_v)
//           [kg 水蒸气/kg 干空气]；p_v 为实际水汽分压。露点模式取
//           p_v = p_ws(Td)（露点即饱和点），相对湿度模式取
//           p_v = RH/100·p_ws(T)。系数 0.621945 为干空气/水蒸气摩尔质量
//           比（ASHRAE Fundamentals 公开公式链 + PsychroLib 语义）。
//           饱和压一律调用族属主 FC_DL_VaporPressureSat，本件零内联公式。
// 开源溯源 (Origin)：改写自 OSCAT Building 行为定义（OSCAT 许可，仅行为定义，零代码行）——道莅 clean-room 实现
// 单位表：T[°C] / Td[°C] / p[Pa] / RH[%] / p_v[Pa] / W[kg 水蒸气/kg 干空气]
// 错误码表：16#0002_2E01 信息级（RH/露点域外已钳位照算，不置 bError）/
//           16#0002_2E10 故障级（大气压非法或输入非有限，置 bError）/
//           16#0002_2E11 故障级（露点>干球等物理矛盾，分母保护，置 bError）/
//           16#0002_2E12 故障级（输入模式枚举非法兜底，置 bError）/
//           16#0002_2E02 预留禁用（不得挪用）
// 状态机：E_DL_RhInputMode（本文件唯一定义，全库唯一属主）：eDewPoint = 0 /
//           eRelativeHumidity = 1；纯计算函数本体无跨拍状态
// 边界行为：① fPress <= 0 → 故障 2E10、bValid := FALSE、W 输出 0；② 任一
//           输入非有限 → 故障 2E10 复用（R90）；③ RH 域外（<0 或 >100）或
//           露点域外（-40~100 °C 外）→ 钳位 + 信息 2E01 + bClamped 照算；
//           ④ p_v >= p（露点 > 干球等物理矛盾）→ 故障 2E11、bValid := FALSE
//           （含湿量分母保护必须故障——与 FC_DL_RhFromDewPoint 的比值钳位
//           策略不同：本件分母直接参与除法，比值件可安全钳 100）；⑤ 枚举
//           非法值走 CASE ELSE 兜底 → 故障 2E12。
// 修订历史：v1.0.0 2026-11-17 首版（R23 派单 · T1-2 焓湿图族拆分②）
//           v1.0.1 2026-11-23 R73 补 bValid 回执：两处 FC_DL_VaporPressureSat
//           调用补收 bValid 局部回执，回执无效并入既有 2E12 兜底分支，契约不变。
//==============================================================================

(*------------------------------------------------------------------------------
 * 枚举: E_DL_RhInputMode（归属本函数，同文件发布，全库唯一定义）
 * 含义: 第二输入 fRhIn 的解释模式，决定 fRhIn 是露点还是相对湿度。
 *-----------------------------------------------------------------------------*)
TYPE E_DL_RhInputMode :
(
    eDewPoint         := 0,  // fRhIn 解释为露点温度 [摄氏度] / fRhIn interpreted as dew-point temperature [degC]
    eRelativeHumidity := 1   // fRhIn 解释为相对湿度 [百分数] / fRhIn interpreted as relative humidity [percent]
);
END_TYPE

(*------------------------------------------------------------------------------
 * 调用示例：bOk := FC_DL_HumidityRatioCalc(fTempC := 25.0,
 *             eRhMode := E_DL_RhInputMode.eRelativeHumidity,
 *             fRhIn := 60.0, fPress := 101325.0,
 *             fHumRatio => fW, fPv => fVp, eErr => uE);
 * 注意：仅当返回 TRUE 且 eErr = 0 时 W 才可进入联锁/能量平衡运算。
 *-----------------------------------------------------------------------------*)
FUNCTION FC_DL_HumidityRatioCalc : BOOL
VAR_INPUT
    fTempC   : LREAL;                    // 干球温度 [摄氏度] / Dry-bulb temperature [degC]
    eRhMode  : E_DL_RhInputMode;         // 第二输入模式枚举 [—] / Interpretation mode of the second input
    fRhIn    : LREAL;                    // 相对湿度 [百分数] 或露点 [摄氏度]，按 eRhMode 解释 / RH [percent] or dew point [degC], per eRhMode
    fPress   : LREAL := 101325.0;        // 大气压 [Pa]，引脚注入非魔法数 / Atmospheric pressure [Pa], injected via the pin
END_VAR
VAR_OUTPUT
    fHumRatio : LREAL;                   // 含湿量 [kg 水蒸气/kg 干空气] / Humidity ratio [kg vapor per kg dry air]
    fPv       : LREAL;                   // 实际水蒸气分压 [Pa] / Actual vapor partial pressure [Pa]
    bClamped  : BOOL;                    // TRUE = 湿度/露点输入已钳位 / TRUE = humidity or dew-point input clamped
    eErr      : UDINT;                   // 错误码，0 = 无错 / Error code, 0 = no error
    bError    : BOOL;                    // 故障级标志，仅故障级错误置位 / Fault-class flag, set only on fault-level codes
    bValid    : BOOL;                    // 输出可用标志 / Outputs usable flag
END_VAR
VAR CONSTANT
    DL_HR_MW_RATIO : LREAL := 0.621945;  // 干空气/水蒸气摩尔质量比 [kg/kg]，ASHRAE 口径 / Molar mass ratio dry air to vapor [kg/kg], ASHRAE
    DL_HR_TD_MIN   : LREAL := -40.0;     // 露点输入钳位下限 [摄氏度]，对齐族属主有效域 / Dew-point clamp floor [degC], aligned with the family owner domain
    DL_HR_TD_MAX   : LREAL := 100.0;     // 露点输入钳位上限 [摄氏度] / Dew-point clamp ceiling [degC]
    DL_HR_RH_MIN   : LREAL := 0.0;       // 相对湿度钳位下限 [百分数] / Relative humidity clamp floor [percent]
    DL_HR_RH_MAX   : LREAL := 100.0;     // 相对湿度钳位上限 [百分数] / Relative humidity clamp ceiling [percent]
    DL_HR_EPS      : LREAL := 1.0E-6;    // 浮点判零容差 [Pa] / Float zero tolerance [Pa]
    DL_HR_INF      : LREAL := 1.7976931348623157E308; // LREAL 幅值上限 / LREAL magnitude ceiling
END_VAR
VAR
    fPwsDb   : LREAL;                    // 干球温度下饱和压 [Pa]，属主件取得 / Saturation pressure at dry bulb [Pa], from the owner FC
    fPwsIn   : LREAL;                    // 第二输入对应饱和压 [Pa] / Saturation pressure of the second input [Pa]
    fRhEff   : LREAL;                    // 钳位后的生效湿度 [百分数] / Effective clamped humidity [percent]
    fTdEff   : LREAL;                    // 钳位后的生效露点 [摄氏度] / Effective clamped dew point [degC]
    fDenom   : LREAL;                    // 含湿量分母 (p − p_v) [Pa] / Humidity ratio denominator [Pa]
    bTdBad   : BOOL;                     // 露点钳位暂存标志 / Staged dew-point clamp flag
    _bPwsValid : BOOL;                   // 饱和压属主件输出可用回执 / Saturation owner FC outputs-usable receipt
    _bPwsClamped : BOOL;    // 属主件钳位回执（本件不消费，仅契约全回执） / Owner clamp receipt (unused, full-receipt contract)
    _nPwsErr     : UDINT;   // 属主件错误码回执 / Owner error-code receipt
    _bPwsError   : BOOL;    // 属主件故障级回执 / Owner fault-flag receipt
END_VAR

(*------------------------------------------------------------------------------
 * 段 1｜出口默认值：入口即赋确定值
 *      Exit defaults: outputs assigned deterministically on entry
 *-----------------------------------------------------------------------------*)
FC_DL_HumidityRatioCalc := FALSE;        // 返回值默认无效 / Return value preset invalid
fHumRatio := 0.0;                        // 含湿量默认置零 / Humidity ratio preset to zero
fPv := 0.0;                              // 水汽分压默认置零 / Vapor pressure preset to zero
bClamped := FALSE;                       // 钳位标志默认 FALSE / Clamped flag preset FALSE
eErr := 16#0000_0000;                    // 错误码先清零 / Error code cleared first
bError := FALSE;                         // 故障标志先清零 / Fault flag cleared first
bValid := FALSE;                         // 可用标志先清零 / Usable flag cleared first
bTdBad := FALSE;                         // 露点钳位暂存清零 / Staged clamp flag cleared

(*------------------------------------------------------------------------------
 * 段 2｜非有限值防御：四个输入全查（含默认注入的大气压）
 *      Non-finite defense on all four inputs including the defaulted pressure
 *-----------------------------------------------------------------------------*)
IF (fTempC <> fTempC) OR (ABS(fTempC) > DL_HR_INF)
   OR (fRhIn <> fRhIn) OR (ABS(fRhIn) > DL_HR_INF)
   OR (fPress <> fPress) OR (ABS(fPress) > DL_HR_INF) THEN
    eErr   := 16#0002_2E10;              // 故障级：输入非有限复用压力非法码（R90） / Fault: non-finite input, code reused
    bError := TRUE;                      // 置故障标志（R45 配对） / Raise the fault flag
    bValid := FALSE;                     // 输出不可用 / Outputs unusable
    RETURN;
END_IF

(*------------------------------------------------------------------------------
 * 段 3｜大气压闸门：p <= 0 物理非法，直接故障（分母保护前置）
 *      Pressure gate: non-positive pressure is physically illegal
 *-----------------------------------------------------------------------------*)
IF fPress <= DL_HR_EPS THEN
    eErr   := 16#0002_2E10;              // 故障级：大气压非法 / Fault: illegal atmospheric pressure
    bError := TRUE;                      // 置故障标志 / Raise the fault flag
    bValid := FALSE;                     // 输出不可用 / Outputs unusable
    RETURN;
END_IF

(*------------------------------------------------------------------------------
 * 段 4｜模式分支：按 eRhMode 解释第二输入，饱和压一律取自族属主件
 *      Mode branch, saturation pressure always from the family owner FC
 *-----------------------------------------------------------------------------*)
CASE eRhMode OF
    E_DL_RhInputMode.eDewPoint:          // 露点模式：p_v = p_ws(Td)，Td 即饱和点
        IF (fRhIn < DL_HR_TD_MIN) OR (fRhIn > DL_HR_TD_MAX) THEN
            fTdEff := MIN(MAX(fRhIn, DL_HR_TD_MIN), DL_HR_TD_MAX); // 露点双侧钳位 / Two-sided dew-point clamp
            bTdBad := TRUE;              // 钳位暂存（信息码在出口统一写，防覆盖） / Staged flag, the info code is written once at the exit
        ELSE
            fTdEff := fRhIn;             // 合法露点原值生效 / Valid dew point applied as-is
        END_IF
        IF (NOT FC_DL_VaporPressureSat(fTempC := fTdEff, fPvSat => fPwsIn, bValid => _bPwsValid, bClamped => _bPwsClamped, eErr => _nPwsErr, bError => _bPwsError)) OR (NOT _bPwsValid) THEN
            eErr   := 16#0002_2E12;      // 故障级：属主件拒绝（其故障即本件故障），兜底码 / Fault: owner FC rejected, fallback code
            bError := TRUE;              // 置故障标志 / Raise the fault flag
            bValid := FALSE;             // 输出不可用 / Outputs unusable
            RETURN;
        END_IF
        fPv := fPwsIn;                   // 露点模式分压 = 露点饱和压 [Pa] / Dew-point mode: partial pressure equals saturation at Td

    E_DL_RhInputMode.eRelativeHumidity:  // 相对湿度模式：p_v = RH/100·p_ws(T)
        IF (fRhIn < DL_HR_RH_MIN) OR (fRhIn > DL_HR_RH_MAX) THEN
            fRhEff := MIN(MAX(fRhIn, DL_HR_RH_MIN), DL_HR_RH_MAX); // 湿度双侧钳位 / Two-sided humidity clamp
            bClamped := TRUE;            // 钳位声明置位 / Clamped flag raised
            eErr := 16#0002_2E01;        // 信息级：RH 已钳位（不置 bError） / Info: RH clamped, no fault flag
        ELSE
            fRhEff := fRhIn;             // 合法湿度原值生效 / Valid humidity applied as-is
        END_IF
        IF (NOT FC_DL_VaporPressureSat(fTempC := fTempC, fPvSat => fPwsDb, bValid => _bPwsValid, bClamped => _bPwsClamped, eErr => _nPwsErr, bError => _bPwsError)) OR (NOT _bPwsValid) THEN
            eErr   := 16#0002_2E12;      // 故障级：属主件拒绝，兜底码 / Fault: owner FC rejected, fallback code
            bError := TRUE;              // 置故障标志 / Raise the fault flag
            bValid := FALSE;             // 输出不可用 / Outputs unusable
            RETURN;
        END_IF
        fPv := (fRhEff / 100.0) * fPwsDb; // 相对湿度模式分压 [Pa] / RH mode partial pressure [Pa]

    ELSE                                 // 枚举非法值兜底（R21：CASE 必带 ELSE）
        eErr   := 16#0002_2E12;          // 故障级：输入模式枚举非法 / Fault: illegal input-mode enum
        bError := TRUE;                  // 置故障标志 / Raise the fault flag
        bValid := FALSE;                 // 输出不可用 / Outputs unusable
        RETURN;
END_CASE

IF bTdBad THEN
    bClamped := TRUE;                    // 露点钳位声明出口统一置位 / Staged dew-point clamp raised at the exit
    eErr := 16#0002_2E01;                // 信息级：露点已钳位（不置 bError） / Info: dew point clamped, no fault flag
END_IF

(*------------------------------------------------------------------------------
 * 段 5｜物理矛盾与分母保护：p_v >= p 或分母过小 → 故障 2E11
 *      Physical contradiction and denominator guard before the division
 *-----------------------------------------------------------------------------*)
fDenom := fPress - fPv;                  // 含湿量分母 [Pa] / Denominator [Pa]
IF (fPv >= fPress) OR (fDenom <= DL_HR_EPS) THEN
    fHumRatio := 0.0;                    // 矛盾输入丢弃，输出确定值 0 / Contradictory input discarded, output zero
    eErr   := 16#0002_2E11;              // 故障级：露点>干球等物理矛盾 / Fault: physical contradiction such as dew point above dry bulb
    bError := TRUE;                      // 置故障标志 / Raise the fault flag
    bValid := FALSE;                     // 输出不可用 / Outputs unusable
    RETURN;
END_IF

(*------------------------------------------------------------------------------
 * 段 6｜含湿量主体：W = 0.621945·p_v/(p − p_v)，分母已闸
 *      Humidity ratio core, denominator already gated
 *-----------------------------------------------------------------------------*)
fHumRatio := DL_HR_MW_RATIO * fPv / fDenom; // 含湿量 [kg 水蒸气/kg 干空气] / Humidity ratio [kg vapor per kg dry air]
bValid := TRUE;                          // 输出可用 / Outputs usable
FC_DL_HumidityRatioCalc := TRUE;         // 返回 TRUE = 计算有效 / Return TRUE = computation valid
END_FUNCTION

(* ---- FC_DL_ZnTune.st ---- *)
(*
  Name        : FC_DL_ZnTune
  Category    : DL_Algo
  Version     : 1.0.0
  Purpose     : Ziegler-Nichols 临界比例度法整定：由临界增益 Ku 与临界振荡周期 Tu 推算 P/PI/PID 三组参数（Kp/Ti/Td 及 Ki/Kd 派生）；/ Ziegler-Nichols ultimate-gain tuning: derive P/PI/PID parameters (Kp, Ti, Td plus Ki, Kd) from Ku and Tu
  溯源        : 借 t2-5-modpid·tune 的分类/参数域组织，clean-room 实现
  Boundary    : ① 组态闸：Ku <= 0 或 Tu <= 0 → 返回 FALSE，全部输出置 0 哨兵（非故障级）；
                ② Ti 派生 Ki 前先判 Ti > eps（P 模式 Ti = 0 → Ki 直接置 0，不做除法）；
                ③ 系数为 ZN 经典表值，属公开表格数据，不含源实现细节；
                ④ 枚举 CASE 含 ELSE 兜底（缺省按 PID 处理，绝不静默输出全零以外的值）。
*)
TYPE E_DL_ZnMode :
(
    eP   := 0,                               (* 纯比例模式 / Pure proportional mode *)
    ePi  := 10,                              (* 比例积分模式 / Proportional-integral mode *)
    ePid := 20                              (* 比例积分微分模式（缺省） / Proportional-integral-derivative mode *)
);
END_TYPE

FUNCTION FC_DL_ZnTune : BOOL
VAR_INPUT
    fKu    : LREAL := 0.0;                   (* 临界增益（等幅振荡时的纯比例增益），域 > 0 [-] / Ultimate gain, must be > 0 *)
    fTu    : LREAL := 0.0;                   (* 临界振荡周期，域 > 0 [s] / Ultimate period, must be > 0 *)
    eMode  : E_DL_ZnMode := E_DL_ZnMode.ePid; (* 整定模式（P/PI/PID）[-] / Tuning mode *)
END_VAR
VAR_OUTPUT
    fKp : LREAL;                             (* 比例增益（无量纲）[-] / Proportional gain *)
    fTi : LREAL;                             (* 积分时间（复位时间），P 模式为 0 [s] / Integral (reset) time, 0 in P mode *)
    fTd : LREAL;                             (* 微分时间（速率时间），P/PI 模式为 0 [s] / Derivative (rate) time, 0 in P/PI *)
    fKi : LREAL;                             (* 积分增益 = Kp / Ti（Ti = 0 时置 0）[1/s] / Integral gain Kp/Ti *)
    fKd : LREAL;                             (* 微分增益 = Kp * Td [s] / Derivative gain Kp*Td *)
END_VAR
VAR CONSTANT
    DL_ZN_EPS    : LREAL := 1.0E-9;          (* 时间量判零容差 [s] / Time epsilon *)
    DL_ZN_KU_P   : LREAL := 0.50;            (* ZN 表：P 模式 Kp = 0.50·Ku [-] / ZN table: P Kp factor *)
    DL_ZN_KU_PI  : LREAL := 0.45;            (* ZN 表：PI 模式 Kp = 0.45·Ku [-] / ZN table: PI Kp factor *)
    DL_ZN_TI_PI  : LREAL := 1.2;             (* ZN 表：PI 模式 Ti = Tu / 1.2 [-] / ZN table: PI Ti divisor *)
    DL_ZN_KU_PID : LREAL := 0.60;            (* ZN 表：PID 模式 Kp = 0.60·Ku [-] / ZN table: PID Kp factor *)
    DL_ZN_TI_PID : LREAL := 2.0;             (* ZN 表：PID 模式 Ti = Tu / 2.0 [-] / ZN table: PID Ti divisor *)
    DL_ZN_TD_PID : LREAL := 8.0;             (* ZN 表：PID 模式 Td = Tu / 8.0 [-] / ZN table: PID Td divisor *)
    DL_ZN_ZERO   : LREAL := 0.0;             (* 零常量（哨兵与占位）[#] / Zero constant *)
END_VAR

(* —— 段 1：输出全路径预置（任何分支都不会留旧值，R191 名实双出口） —— *)
fKp := DL_ZN_ZERO;                           (* Kp 预置 0 / Kp preset *)
fTi := DL_ZN_ZERO;                           (* Ti 预置 0 / Ti preset *)
fTd := DL_ZN_ZERO;                           (* Td 预置 0 / Td preset *)
fKi := DL_ZN_ZERO;                           (* Ki 预置 0 / Ki preset *)
fKd := DL_ZN_ZERO;                           (* Kd 预置 0 / Kd preset *)
FC_DL_ZnTune := FALSE;                       (* 返回值预置 FALSE：仅合法分支翻 TRUE / Return preset FALSE *)

(* —— 段 2：非有限输入拒收（NaN 自反 + Inf 差判） —— *)
IF (fKu <> fKu) OR (fTu <> fTu) THEN
    RETURN;                                  (* NaN 拒收 / NaN rejected *)
END_IF
IF ((fKu - fKu) <> (fKu - fKu)) OR ((fTu - fTu) <> (fTu - fTu)) THEN
    RETURN;                                  (* Inf 拒收 / Inf rejected *)
END_IF

(* —— 段 3：组态闸（Ku/Tu 正域，除子唯一出入口） —— *)
IF (fKu <= DL_ZN_EPS) OR (fTu <= DL_ZN_EPS) THEN
    RETURN;                                  (* 临界参数非正：无整定语义，返回 FALSE + 零哨兵 / Non-positive Ku/Tu: sentinel *)
END_IF

(* —— 段 4：按模式取 ZN 表系数（CASE 含 ELSE 兜底为 PID） —— *)
CASE eMode OF
    E_DL_ZnMode.eP:                          (* P 模式：仅 Kp，Ti/Td 保持 0 / P mode *)
        fKp := DL_ZN_KU_P * fKu;             (* Kp = 0.50·Ku [-] / Kp *)
    E_DL_ZnMode.ePi:                         (* PI 模式：Kp + Ti / PI mode *)
        fKp := DL_ZN_KU_PI * fKu;            (* Kp = 0.45·Ku [-] / Kp *)
        fTi := fTu / DL_ZN_TI_PI;            (* Ti = Tu/1.2，除子为表常量非 0 [s] / Ti *)
    E_DL_ZnMode.ePid:                        (* PID 模式：Kp + Ti + Td / PID mode *)
        fKp := DL_ZN_KU_PID * fKu;           (* Kp = 0.60·Ku [-] / Kp *)
        fTi := fTu / DL_ZN_TI_PID;           (* Ti = Tu/2.0 [s] / Ti *)
        fTd := fTu / DL_ZN_TD_PID;           (* Td = Tu/8.0 [s] / Td *)
    ELSE                                     (* 非法模式：按 PID 兜底，不静默清零 / Illegal mode: fallback to PID *)
        fKp := DL_ZN_KU_PID * fKu;           (* 兜底 Kp = 0.60·Ku [-] / Fallback Kp *)
        fTi := fTu / DL_ZN_TI_PID;           (* 兜底 Ti [s] / Fallback Ti *)
        fTd := fTu / DL_ZN_TD_PID;           (* 兜底 Td [s] / Fallback Td *)
END_CASE

(* —— 段 5：Ki/Kd 派生（Ti 判零后再除，P 模式 Ki 保持 0） —— *)
IF ABS(fTi) > DL_ZN_EPS THEN
    fKi := fKp / fTi;                        (* Ki = Kp/Ti，除子已过容差闸 [1/s] / Ki, divisor gated *)
ELSE
    fKi := DL_ZN_ZERO;                       (* Ti = 0：积分增益无定义，置 0 / Ti zero: Ki 0 *)
END_IF
fKd := fKp * fTd;                            (* Kd = Kp·Td（乘性派生无除零）[s] / Kd, multiplicative *)
FC_DL_ZnTune := TRUE;                        (* 参数全套有效 / All parameters valid *)
END_FUNCTION
